(* IEC 61131-3 sources: STAR-PLC-Agent/results/raw/codex_matrix_resume_20261114/codex_deepseek/PUB011/functional/attempt_0001, 1 file *)

(* ---- test_program.st ---- *)
PROGRAM PLC_PRG
VAR
 BenchStep : UDINT := 0;
 BenchCalls : UDINT := 0;
 BenchDone : BOOL := FALSE;
 BenchUut0 : FB_Task;
 BenchUut1 : FB_Task;
 BenchUut2 : FB_Task;
 BenchUut3 : FB_Task;
 BenchUut4 : FB_Task;
 BenchUut5 : FB_Task;
 BenchUut6 : FB_Task;
 BenchUut7 : FB_Task;
 TraceIn_Mode : ARRAY[0..81] OF BOOL;
 TraceIn_ForwardButton : ARRAY[0..81] OF BOOL;
 TraceIn_ReverseButton : ARRAY[0..81] OF BOOL;
 TraceIn_SensorA : ARRAY[0..81] OF BOOL;
 TraceIn_SensorB : ARRAY[0..81] OF BOOL;
 TraceIn_SensorC : ARRAY[0..81] OF BOOL;
 TraceIn_ButtonA : ARRAY[0..81] OF BOOL;
 TraceIn_ButtonB : ARRAY[0..81] OF BOOL;
 TraceIn_ButtonC : ARRAY[0..81] OF BOOL;
 TraceOut_MotorForward : ARRAY[0..81] OF BOOL;
 TraceOut_MotorReverse : ARRAY[0..81] OF BOOL;
 TraceOut_CompletionLight : ARRAY[0..81] OF BOOL;
END_VAR

IF NOT BenchDone THEN
 CASE BenchStep OF
 0:
   BenchUut0.Mode := FALSE;
   BenchUut0.ForwardButton := FALSE;
   BenchUut0.ReverseButton := FALSE;
   BenchUut0.SensorA := FALSE;
   BenchUut0.SensorB := FALSE;
   BenchUut0.SensorC := FALSE;
   BenchUut0.ButtonA := FALSE;
   BenchUut0.ButtonB := FALSE;
   BenchUut0.ButtonC := FALSE;
   TraceIn_Mode[0] := BenchUut0.Mode;
   TraceIn_ForwardButton[0] := BenchUut0.ForwardButton;
   TraceIn_ReverseButton[0] := BenchUut0.ReverseButton;
   TraceIn_SensorA[0] := BenchUut0.SensorA;
   TraceIn_SensorB[0] := BenchUut0.SensorB;
   TraceIn_SensorC[0] := BenchUut0.SensorC;
   TraceIn_ButtonA[0] := BenchUut0.ButtonA;
   TraceIn_ButtonB[0] := BenchUut0.ButtonB;
   TraceIn_ButtonC[0] := BenchUut0.ButtonC;
   BenchUut0();
   TraceOut_MotorForward[0] := BenchUut0.MotorForward;
   TraceOut_MotorReverse[0] := BenchUut0.MotorReverse;
   TraceOut_CompletionLight[0] := BenchUut0.CompletionLight;
   BenchCalls := BenchCalls + 1;
 1:
   BenchUut0.Mode := FALSE;
   BenchUut0.ForwardButton := TRUE;
   BenchUut0.ReverseButton := FALSE;
   BenchUut0.SensorA := FALSE;
   BenchUut0.SensorB := FALSE;
   BenchUut0.SensorC := FALSE;
   BenchUut0.ButtonA := FALSE;
   BenchUut0.ButtonB := FALSE;
   BenchUut0.ButtonC := FALSE;
   TraceIn_Mode[1] := BenchUut0.Mode;
   TraceIn_ForwardButton[1] := BenchUut0.ForwardButton;
   TraceIn_ReverseButton[1] := BenchUut0.ReverseButton;
   TraceIn_SensorA[1] := BenchUut0.SensorA;
   TraceIn_SensorB[1] := BenchUut0.SensorB;
   TraceIn_SensorC[1] := BenchUut0.SensorC;
   TraceIn_ButtonA[1] := BenchUut0.ButtonA;
   TraceIn_ButtonB[1] := BenchUut0.ButtonB;
   TraceIn_ButtonC[1] := BenchUut0.ButtonC;
   BenchUut0();
   TraceOut_MotorForward[1] := BenchUut0.MotorForward;
   TraceOut_MotorReverse[1] := BenchUut0.MotorReverse;
   TraceOut_CompletionLight[1] := BenchUut0.CompletionLight;
   BenchCalls := BenchCalls + 1;
 2:
   BenchUut0.Mode := FALSE;
   BenchUut0.ForwardButton := FALSE;
   BenchUut0.ReverseButton := TRUE;
   BenchUut0.SensorA := FALSE;
   BenchUut0.SensorB := FALSE;
   BenchUut0.SensorC := FALSE;
   BenchUut0.ButtonA := FALSE;
   BenchUut0.ButtonB := FALSE;
   BenchUut0.ButtonC := FALSE;
   TraceIn_Mode[2] := BenchUut0.Mode;
   TraceIn_ForwardButton[2] := BenchUut0.ForwardButton;
   TraceIn_ReverseButton[2] := BenchUut0.ReverseButton;
   TraceIn_SensorA[2] := BenchUut0.SensorA;
   TraceIn_SensorB[2] := BenchUut0.SensorB;
   TraceIn_SensorC[2] := BenchUut0.SensorC;
   TraceIn_ButtonA[2] := BenchUut0.ButtonA;
   TraceIn_ButtonB[2] := BenchUut0.ButtonB;
   TraceIn_ButtonC[2] := BenchUut0.ButtonC;
   BenchUut0();
   TraceOut_MotorForward[2] := BenchUut0.MotorForward;
   TraceOut_MotorReverse[2] := BenchUut0.MotorReverse;
   TraceOut_CompletionLight[2] := BenchUut0.CompletionLight;
   BenchCalls := BenchCalls + 1;
 3:
   BenchUut1.Mode := TRUE;
   BenchUut1.ForwardButton := FALSE;
   BenchUut1.ReverseButton := FALSE;
   BenchUut1.SensorA := FALSE;
   BenchUut1.SensorB := FALSE;
   BenchUut1.SensorC := FALSE;
   BenchUut1.ButtonA := FALSE;
   BenchUut1.ButtonB := FALSE;
   BenchUut1.ButtonC := FALSE;
   TraceIn_Mode[3] := BenchUut1.Mode;
   TraceIn_ForwardButton[3] := BenchUut1.ForwardButton;
   TraceIn_ReverseButton[3] := BenchUut1.ReverseButton;
   TraceIn_SensorA[3] := BenchUut1.SensorA;
   TraceIn_SensorB[3] := BenchUut1.SensorB;
   TraceIn_SensorC[3] := BenchUut1.SensorC;
   TraceIn_ButtonA[3] := BenchUut1.ButtonA;
   TraceIn_ButtonB[3] := BenchUut1.ButtonB;
   TraceIn_ButtonC[3] := BenchUut1.ButtonC;
   BenchUut1();
   TraceOut_MotorForward[3] := BenchUut1.MotorForward;
   TraceOut_MotorReverse[3] := BenchUut1.MotorReverse;
   TraceOut_CompletionLight[3] := BenchUut1.CompletionLight;
   BenchCalls := BenchCalls + 1;
 4:
   BenchUut1.Mode := TRUE;
   BenchUut1.ForwardButton := FALSE;
   BenchUut1.ReverseButton := FALSE;
   BenchUut1.SensorA := TRUE;
   BenchUut1.SensorB := FALSE;
   BenchUut1.SensorC := FALSE;
   BenchUut1.ButtonA := FALSE;
   BenchUut1.ButtonB := FALSE;
   BenchUut1.ButtonC := FALSE;
   TraceIn_Mode[4] := BenchUut1.Mode;
   TraceIn_ForwardButton[4] := BenchUut1.ForwardButton;
   TraceIn_ReverseButton[4] := BenchUut1.ReverseButton;
   TraceIn_SensorA[4] := BenchUut1.SensorA;
   TraceIn_SensorB[4] := BenchUut1.SensorB;
   TraceIn_SensorC[4] := BenchUut1.SensorC;
   TraceIn_ButtonA[4] := BenchUut1.ButtonA;
   TraceIn_ButtonB[4] := BenchUut1.ButtonB;
   TraceIn_ButtonC[4] := BenchUut1.ButtonC;
   BenchUut1();
   TraceOut_MotorForward[4] := BenchUut1.MotorForward;
   TraceOut_MotorReverse[4] := BenchUut1.MotorReverse;
   TraceOut_CompletionLight[4] := BenchUut1.CompletionLight;
   BenchCalls := BenchCalls + 1;
 5:
   BenchUut1.Mode := TRUE;
   BenchUut1.ForwardButton := FALSE;
   BenchUut1.ReverseButton := FALSE;
   BenchUut1.SensorA := TRUE;
   BenchUut1.SensorB := FALSE;
   BenchUut1.SensorC := FALSE;
   BenchUut1.ButtonA := TRUE;
   BenchUut1.ButtonB := FALSE;
   BenchUut1.ButtonC := FALSE;
   TraceIn_Mode[5] := BenchUut1.Mode;
   TraceIn_ForwardButton[5] := BenchUut1.ForwardButton;
   TraceIn_ReverseButton[5] := BenchUut1.ReverseButton;
   TraceIn_SensorA[5] := BenchUut1.SensorA;
   TraceIn_SensorB[5] := BenchUut1.SensorB;
   TraceIn_SensorC[5] := BenchUut1.SensorC;
   TraceIn_ButtonA[5] := BenchUut1.ButtonA;
   TraceIn_ButtonB[5] := BenchUut1.ButtonB;
   TraceIn_ButtonC[5] := BenchUut1.ButtonC;
   BenchUut1();
   TraceOut_MotorForward[5] := BenchUut1.MotorForward;
   TraceOut_MotorReverse[5] := BenchUut1.MotorReverse;
   TraceOut_CompletionLight[5] := BenchUut1.CompletionLight;
   BenchCalls := BenchCalls + 1;
 6:
   BenchUut1.Mode := TRUE;
   BenchUut1.ForwardButton := FALSE;
   BenchUut1.ReverseButton := FALSE;
   BenchUut1.SensorA := FALSE;
   BenchUut1.SensorB := FALSE;
   BenchUut1.SensorC := FALSE;
   BenchUut1.ButtonA := FALSE;
   BenchUut1.ButtonB := FALSE;
   BenchUut1.ButtonC := FALSE;
   TraceIn_Mode[6] := BenchUut1.Mode;
   TraceIn_ForwardButton[6] := BenchUut1.ForwardButton;
   TraceIn_ReverseButton[6] := BenchUut1.ReverseButton;
   TraceIn_SensorA[6] := BenchUut1.SensorA;
   TraceIn_SensorB[6] := BenchUut1.SensorB;
   TraceIn_SensorC[6] := BenchUut1.SensorC;
   TraceIn_ButtonA[6] := BenchUut1.ButtonA;
   TraceIn_ButtonB[6] := BenchUut1.ButtonB;
   TraceIn_ButtonC[6] := BenchUut1.ButtonC;
   BenchUut1();
   TraceOut_MotorForward[6] := BenchUut1.MotorForward;
   TraceOut_MotorReverse[6] := BenchUut1.MotorReverse;
   TraceOut_CompletionLight[6] := BenchUut1.CompletionLight;
   BenchCalls := BenchCalls + 1;
 7:
   BenchUut1.Mode := TRUE;
   BenchUut1.ForwardButton := FALSE;
   BenchUut1.ReverseButton := FALSE;
   BenchUut1.SensorA := FALSE;
   BenchUut1.SensorB := TRUE;
   BenchUut1.SensorC := FALSE;
   BenchUut1.ButtonA := FALSE;
   BenchUut1.ButtonB := FALSE;
   BenchUut1.ButtonC := FALSE;
   TraceIn_Mode[7] := BenchUut1.Mode;
   TraceIn_ForwardButton[7] := BenchUut1.ForwardButton;
   TraceIn_ReverseButton[7] := BenchUut1.ReverseButton;
   TraceIn_SensorA[7] := BenchUut1.SensorA;
   TraceIn_SensorB[7] := BenchUut1.SensorB;
   TraceIn_SensorC[7] := BenchUut1.SensorC;
   TraceIn_ButtonA[7] := BenchUut1.ButtonA;
   TraceIn_ButtonB[7] := BenchUut1.ButtonB;
   TraceIn_ButtonC[7] := BenchUut1.ButtonC;
   BenchUut1();
   TraceOut_MotorForward[7] := BenchUut1.MotorForward;
   TraceOut_MotorReverse[7] := BenchUut1.MotorReverse;
   TraceOut_CompletionLight[7] := BenchUut1.CompletionLight;
   BenchCalls := BenchCalls + 1;
 8:
   BenchUut1.Mode := TRUE;
   BenchUut1.ForwardButton := FALSE;
   BenchUut1.ReverseButton := FALSE;
   BenchUut1.SensorA := FALSE;
   BenchUut1.SensorB := TRUE;
   BenchUut1.SensorC := FALSE;
   BenchUut1.ButtonA := FALSE;
   BenchUut1.ButtonB := TRUE;
   BenchUut1.ButtonC := FALSE;
   TraceIn_Mode[8] := BenchUut1.Mode;
   TraceIn_ForwardButton[8] := BenchUut1.ForwardButton;
   TraceIn_ReverseButton[8] := BenchUut1.ReverseButton;
   TraceIn_SensorA[8] := BenchUut1.SensorA;
   TraceIn_SensorB[8] := BenchUut1.SensorB;
   TraceIn_SensorC[8] := BenchUut1.SensorC;
   TraceIn_ButtonA[8] := BenchUut1.ButtonA;
   TraceIn_ButtonB[8] := BenchUut1.ButtonB;
   TraceIn_ButtonC[8] := BenchUut1.ButtonC;
   BenchUut1();
   TraceOut_MotorForward[8] := BenchUut1.MotorForward;
   TraceOut_MotorReverse[8] := BenchUut1.MotorReverse;
   TraceOut_CompletionLight[8] := BenchUut1.CompletionLight;
   BenchCalls := BenchCalls + 1;
 9:
   BenchUut1.Mode := TRUE;
   BenchUut1.ForwardButton := FALSE;
   BenchUut1.ReverseButton := FALSE;
   BenchUut1.SensorA := FALSE;
   BenchUut1.SensorB := FALSE;
   BenchUut1.SensorC := TRUE;
   BenchUut1.ButtonA := FALSE;
   BenchUut1.ButtonB := FALSE;
   BenchUut1.ButtonC := FALSE;
   TraceIn_Mode[9] := BenchUut1.Mode;
   TraceIn_ForwardButton[9] := BenchUut1.ForwardButton;
   TraceIn_ReverseButton[9] := BenchUut1.ReverseButton;
   TraceIn_SensorA[9] := BenchUut1.SensorA;
   TraceIn_SensorB[9] := BenchUut1.SensorB;
   TraceIn_SensorC[9] := BenchUut1.SensorC;
   TraceIn_ButtonA[9] := BenchUut1.ButtonA;
   TraceIn_ButtonB[9] := BenchUut1.ButtonB;
   TraceIn_ButtonC[9] := BenchUut1.ButtonC;
   BenchUut1();
   TraceOut_MotorForward[9] := BenchUut1.MotorForward;
   TraceOut_MotorReverse[9] := BenchUut1.MotorReverse;
   TraceOut_CompletionLight[9] := BenchUut1.CompletionLight;
   BenchCalls := BenchCalls + 1;
 10:
   BenchUut1.Mode := TRUE;
   BenchUut1.ForwardButton := FALSE;
   BenchUut1.ReverseButton := FALSE;
   BenchUut1.SensorA := FALSE;
   BenchUut1.SensorB := FALSE;
   BenchUut1.SensorC := TRUE;
   BenchUut1.ButtonA := FALSE;
   BenchUut1.ButtonB := FALSE;
   BenchUut1.ButtonC := TRUE;
   TraceIn_Mode[10] := BenchUut1.Mode;
   TraceIn_ForwardButton[10] := BenchUut1.ForwardButton;
   TraceIn_ReverseButton[10] := BenchUut1.ReverseButton;
   TraceIn_SensorA[10] := BenchUut1.SensorA;
   TraceIn_SensorB[10] := BenchUut1.SensorB;
   TraceIn_SensorC[10] := BenchUut1.SensorC;
   TraceIn_ButtonA[10] := BenchUut1.ButtonA;
   TraceIn_ButtonB[10] := BenchUut1.ButtonB;
   TraceIn_ButtonC[10] := BenchUut1.ButtonC;
   BenchUut1();
   TraceOut_MotorForward[10] := BenchUut1.MotorForward;
   TraceOut_MotorReverse[10] := BenchUut1.MotorReverse;
   TraceOut_CompletionLight[10] := BenchUut1.CompletionLight;
   BenchCalls := BenchCalls + 1;
 11:
   BenchUut1.Mode := TRUE;
   BenchUut1.ForwardButton := FALSE;
   BenchUut1.ReverseButton := FALSE;
   BenchUut1.SensorA := FALSE;
   BenchUut1.SensorB := FALSE;
   BenchUut1.SensorC := TRUE;
   BenchUut1.ButtonA := FALSE;
   BenchUut1.ButtonB := FALSE;
   BenchUut1.ButtonC := FALSE;
   TraceIn_Mode[11] := BenchUut1.Mode;
   TraceIn_ForwardButton[11] := BenchUut1.ForwardButton;
   TraceIn_ReverseButton[11] := BenchUut1.ReverseButton;
   TraceIn_SensorA[11] := BenchUut1.SensorA;
   TraceIn_SensorB[11] := BenchUut1.SensorB;
   TraceIn_SensorC[11] := BenchUut1.SensorC;
   TraceIn_ButtonA[11] := BenchUut1.ButtonA;
   TraceIn_ButtonB[11] := BenchUut1.ButtonB;
   TraceIn_ButtonC[11] := BenchUut1.ButtonC;
   BenchUut1();
   TraceOut_MotorForward[11] := BenchUut1.MotorForward;
   TraceOut_MotorReverse[11] := BenchUut1.MotorReverse;
   TraceOut_CompletionLight[11] := BenchUut1.CompletionLight;
   BenchCalls := BenchCalls + 1;
 12:
   BenchUut1.Mode := TRUE;
   BenchUut1.ForwardButton := FALSE;
   BenchUut1.ReverseButton := FALSE;
   BenchUut1.SensorA := FALSE;
   BenchUut1.SensorB := FALSE;
   BenchUut1.SensorC := FALSE;
   BenchUut1.ButtonA := FALSE;
   BenchUut1.ButtonB := FALSE;
   BenchUut1.ButtonC := FALSE;
   TraceIn_Mode[12] := BenchUut1.Mode;
   TraceIn_ForwardButton[12] := BenchUut1.ForwardButton;
   TraceIn_ReverseButton[12] := BenchUut1.ReverseButton;
   TraceIn_SensorA[12] := BenchUut1.SensorA;
   TraceIn_SensorB[12] := BenchUut1.SensorB;
   TraceIn_SensorC[12] := BenchUut1.SensorC;
   TraceIn_ButtonA[12] := BenchUut1.ButtonA;
   TraceIn_ButtonB[12] := BenchUut1.ButtonB;
   TraceIn_ButtonC[12] := BenchUut1.ButtonC;
   BenchUut1();
   TraceOut_MotorForward[12] := BenchUut1.MotorForward;
   TraceOut_MotorReverse[12] := BenchUut1.MotorReverse;
   TraceOut_CompletionLight[12] := BenchUut1.CompletionLight;
   BenchCalls := BenchCalls + 1;
 13:
   BenchUut2.Mode := TRUE;
   BenchUut2.ForwardButton := FALSE;
   BenchUut2.ReverseButton := FALSE;
   BenchUut2.SensorA := FALSE;
   BenchUut2.SensorB := FALSE;
   BenchUut2.SensorC := FALSE;
   BenchUut2.ButtonA := FALSE;
   BenchUut2.ButtonB := TRUE;
   BenchUut2.ButtonC := TRUE;
   TraceIn_Mode[13] := BenchUut2.Mode;
   TraceIn_ForwardButton[13] := BenchUut2.ForwardButton;
   TraceIn_ReverseButton[13] := BenchUut2.ReverseButton;
   TraceIn_SensorA[13] := BenchUut2.SensorA;
   TraceIn_SensorB[13] := BenchUut2.SensorB;
   TraceIn_SensorC[13] := BenchUut2.SensorC;
   TraceIn_ButtonA[13] := BenchUut2.ButtonA;
   TraceIn_ButtonB[13] := BenchUut2.ButtonB;
   TraceIn_ButtonC[13] := BenchUut2.ButtonC;
   BenchUut2();
   TraceOut_MotorForward[13] := BenchUut2.MotorForward;
   TraceOut_MotorReverse[13] := BenchUut2.MotorReverse;
   TraceOut_CompletionLight[13] := BenchUut2.CompletionLight;
   BenchCalls := BenchCalls + 1;
 14:
   BenchUut2.Mode := TRUE;
   BenchUut2.ForwardButton := FALSE;
   BenchUut2.ReverseButton := FALSE;
   BenchUut2.SensorA := TRUE;
   BenchUut2.SensorB := FALSE;
   BenchUut2.SensorC := FALSE;
   BenchUut2.ButtonA := FALSE;
   BenchUut2.ButtonB := TRUE;
   BenchUut2.ButtonC := FALSE;
   TraceIn_Mode[14] := BenchUut2.Mode;
   TraceIn_ForwardButton[14] := BenchUut2.ForwardButton;
   TraceIn_ReverseButton[14] := BenchUut2.ReverseButton;
   TraceIn_SensorA[14] := BenchUut2.SensorA;
   TraceIn_SensorB[14] := BenchUut2.SensorB;
   TraceIn_SensorC[14] := BenchUut2.SensorC;
   TraceIn_ButtonA[14] := BenchUut2.ButtonA;
   TraceIn_ButtonB[14] := BenchUut2.ButtonB;
   TraceIn_ButtonC[14] := BenchUut2.ButtonC;
   BenchUut2();
   TraceOut_MotorForward[14] := BenchUut2.MotorForward;
   TraceOut_MotorReverse[14] := BenchUut2.MotorReverse;
   TraceOut_CompletionLight[14] := BenchUut2.CompletionLight;
   BenchCalls := BenchCalls + 1;
 15:
   BenchUut3.Mode := TRUE;
   BenchUut3.ForwardButton := FALSE;
   BenchUut3.ReverseButton := FALSE;
   BenchUut3.SensorA := FALSE;
   BenchUut3.SensorB := FALSE;
   BenchUut3.SensorC := FALSE;
   BenchUut3.ButtonA := FALSE;
   BenchUut3.ButtonB := FALSE;
   BenchUut3.ButtonC := FALSE;
   TraceIn_Mode[15] := BenchUut3.Mode;
   TraceIn_ForwardButton[15] := BenchUut3.ForwardButton;
   TraceIn_ReverseButton[15] := BenchUut3.ReverseButton;
   TraceIn_SensorA[15] := BenchUut3.SensorA;
   TraceIn_SensorB[15] := BenchUut3.SensorB;
   TraceIn_SensorC[15] := BenchUut3.SensorC;
   TraceIn_ButtonA[15] := BenchUut3.ButtonA;
   TraceIn_ButtonB[15] := BenchUut3.ButtonB;
   TraceIn_ButtonC[15] := BenchUut3.ButtonC;
   BenchUut3();
   TraceOut_MotorForward[15] := BenchUut3.MotorForward;
   TraceOut_MotorReverse[15] := BenchUut3.MotorReverse;
   TraceOut_CompletionLight[15] := BenchUut3.CompletionLight;
   BenchCalls := BenchCalls + 1;
 16:
   BenchUut3.Mode := TRUE;
   BenchUut3.ForwardButton := FALSE;
   BenchUut3.ReverseButton := FALSE;
   BenchUut3.SensorA := TRUE;
   BenchUut3.SensorB := FALSE;
   BenchUut3.SensorC := FALSE;
   BenchUut3.ButtonA := FALSE;
   BenchUut3.ButtonB := FALSE;
   BenchUut3.ButtonC := FALSE;
   TraceIn_Mode[16] := BenchUut3.Mode;
   TraceIn_ForwardButton[16] := BenchUut3.ForwardButton;
   TraceIn_ReverseButton[16] := BenchUut3.ReverseButton;
   TraceIn_SensorA[16] := BenchUut3.SensorA;
   TraceIn_SensorB[16] := BenchUut3.SensorB;
   TraceIn_SensorC[16] := BenchUut3.SensorC;
   TraceIn_ButtonA[16] := BenchUut3.ButtonA;
   TraceIn_ButtonB[16] := BenchUut3.ButtonB;
   TraceIn_ButtonC[16] := BenchUut3.ButtonC;
   BenchUut3();
   TraceOut_MotorForward[16] := BenchUut3.MotorForward;
   TraceOut_MotorReverse[16] := BenchUut3.MotorReverse;
   TraceOut_CompletionLight[16] := BenchUut3.CompletionLight;
   BenchCalls := BenchCalls + 1;
 17:
   BenchUut3.Mode := TRUE;
   BenchUut3.ForwardButton := FALSE;
   BenchUut3.ReverseButton := FALSE;
   BenchUut3.SensorA := TRUE;
   BenchUut3.SensorB := FALSE;
   BenchUut3.SensorC := FALSE;
   BenchUut3.ButtonA := TRUE;
   BenchUut3.ButtonB := FALSE;
   BenchUut3.ButtonC := FALSE;
   TraceIn_Mode[17] := BenchUut3.Mode;
   TraceIn_ForwardButton[17] := BenchUut3.ForwardButton;
   TraceIn_ReverseButton[17] := BenchUut3.ReverseButton;
   TraceIn_SensorA[17] := BenchUut3.SensorA;
   TraceIn_SensorB[17] := BenchUut3.SensorB;
   TraceIn_SensorC[17] := BenchUut3.SensorC;
   TraceIn_ButtonA[17] := BenchUut3.ButtonA;
   TraceIn_ButtonB[17] := BenchUut3.ButtonB;
   TraceIn_ButtonC[17] := BenchUut3.ButtonC;
   BenchUut3();
   TraceOut_MotorForward[17] := BenchUut3.MotorForward;
   TraceOut_MotorReverse[17] := BenchUut3.MotorReverse;
   TraceOut_CompletionLight[17] := BenchUut3.CompletionLight;
   BenchCalls := BenchCalls + 1;
 18:
   BenchUut3.Mode := TRUE;
   BenchUut3.ForwardButton := FALSE;
   BenchUut3.ReverseButton := FALSE;
   BenchUut3.SensorA := FALSE;
   BenchUut3.SensorB := FALSE;
   BenchUut3.SensorC := FALSE;
   BenchUut3.ButtonA := FALSE;
   BenchUut3.ButtonB := FALSE;
   BenchUut3.ButtonC := FALSE;
   TraceIn_Mode[18] := BenchUut3.Mode;
   TraceIn_ForwardButton[18] := BenchUut3.ForwardButton;
   TraceIn_ReverseButton[18] := BenchUut3.ReverseButton;
   TraceIn_SensorA[18] := BenchUut3.SensorA;
   TraceIn_SensorB[18] := BenchUut3.SensorB;
   TraceIn_SensorC[18] := BenchUut3.SensorC;
   TraceIn_ButtonA[18] := BenchUut3.ButtonA;
   TraceIn_ButtonB[18] := BenchUut3.ButtonB;
   TraceIn_ButtonC[18] := BenchUut3.ButtonC;
   BenchUut3();
   TraceOut_MotorForward[18] := BenchUut3.MotorForward;
   TraceOut_MotorReverse[18] := BenchUut3.MotorReverse;
   TraceOut_CompletionLight[18] := BenchUut3.CompletionLight;
   BenchCalls := BenchCalls + 1;
 19:
   BenchUut3.Mode := TRUE;
   BenchUut3.ForwardButton := FALSE;
   BenchUut3.ReverseButton := FALSE;
   BenchUut3.SensorA := FALSE;
   BenchUut3.SensorB := TRUE;
   BenchUut3.SensorC := FALSE;
   BenchUut3.ButtonA := FALSE;
   BenchUut3.ButtonB := FALSE;
   BenchUut3.ButtonC := FALSE;
   TraceIn_Mode[19] := BenchUut3.Mode;
   TraceIn_ForwardButton[19] := BenchUut3.ForwardButton;
   TraceIn_ReverseButton[19] := BenchUut3.ReverseButton;
   TraceIn_SensorA[19] := BenchUut3.SensorA;
   TraceIn_SensorB[19] := BenchUut3.SensorB;
   TraceIn_SensorC[19] := BenchUut3.SensorC;
   TraceIn_ButtonA[19] := BenchUut3.ButtonA;
   TraceIn_ButtonB[19] := BenchUut3.ButtonB;
   TraceIn_ButtonC[19] := BenchUut3.ButtonC;
   BenchUut3();
   TraceOut_MotorForward[19] := BenchUut3.MotorForward;
   TraceOut_MotorReverse[19] := BenchUut3.MotorReverse;
   TraceOut_CompletionLight[19] := BenchUut3.CompletionLight;
   BenchCalls := BenchCalls + 1;
 20:
   BenchUut3.Mode := TRUE;
   BenchUut3.ForwardButton := FALSE;
   BenchUut3.ReverseButton := FALSE;
   BenchUut3.SensorA := FALSE;
   BenchUut3.SensorB := TRUE;
   BenchUut3.SensorC := FALSE;
   BenchUut3.ButtonA := FALSE;
   BenchUut3.ButtonB := TRUE;
   BenchUut3.ButtonC := FALSE;
   TraceIn_Mode[20] := BenchUut3.Mode;
   TraceIn_ForwardButton[20] := BenchUut3.ForwardButton;
   TraceIn_ReverseButton[20] := BenchUut3.ReverseButton;
   TraceIn_SensorA[20] := BenchUut3.SensorA;
   TraceIn_SensorB[20] := BenchUut3.SensorB;
   TraceIn_SensorC[20] := BenchUut3.SensorC;
   TraceIn_ButtonA[20] := BenchUut3.ButtonA;
   TraceIn_ButtonB[20] := BenchUut3.ButtonB;
   TraceIn_ButtonC[20] := BenchUut3.ButtonC;
   BenchUut3();
   TraceOut_MotorForward[20] := BenchUut3.MotorForward;
   TraceOut_MotorReverse[20] := BenchUut3.MotorReverse;
   TraceOut_CompletionLight[20] := BenchUut3.CompletionLight;
   BenchCalls := BenchCalls + 1;
 21:
   BenchUut3.Mode := TRUE;
   BenchUut3.ForwardButton := FALSE;
   BenchUut3.ReverseButton := FALSE;
   BenchUut3.SensorA := FALSE;
   BenchUut3.SensorB := FALSE;
   BenchUut3.SensorC := FALSE;
   BenchUut3.ButtonA := FALSE;
   BenchUut3.ButtonB := FALSE;
   BenchUut3.ButtonC := FALSE;
   TraceIn_Mode[21] := BenchUut3.Mode;
   TraceIn_ForwardButton[21] := BenchUut3.ForwardButton;
   TraceIn_ReverseButton[21] := BenchUut3.ReverseButton;
   TraceIn_SensorA[21] := BenchUut3.SensorA;
   TraceIn_SensorB[21] := BenchUut3.SensorB;
   TraceIn_SensorC[21] := BenchUut3.SensorC;
   TraceIn_ButtonA[21] := BenchUut3.ButtonA;
   TraceIn_ButtonB[21] := BenchUut3.ButtonB;
   TraceIn_ButtonC[21] := BenchUut3.ButtonC;
   BenchUut3();
   TraceOut_MotorForward[21] := BenchUut3.MotorForward;
   TraceOut_MotorReverse[21] := BenchUut3.MotorReverse;
   TraceOut_CompletionLight[21] := BenchUut3.CompletionLight;
   BenchCalls := BenchCalls + 1;
 22:
   BenchUut4.Mode := TRUE;
   BenchUut4.ForwardButton := FALSE;
   BenchUut4.ReverseButton := FALSE;
   BenchUut4.SensorA := TRUE;
   BenchUut4.SensorB := FALSE;
   BenchUut4.SensorC := FALSE;
   BenchUut4.ButtonA := TRUE;
   BenchUut4.ButtonB := FALSE;
   BenchUut4.ButtonC := FALSE;
   TraceIn_Mode[22] := BenchUut4.Mode;
   TraceIn_ForwardButton[22] := BenchUut4.ForwardButton;
   TraceIn_ReverseButton[22] := BenchUut4.ReverseButton;
   TraceIn_SensorA[22] := BenchUut4.SensorA;
   TraceIn_SensorB[22] := BenchUut4.SensorB;
   TraceIn_SensorC[22] := BenchUut4.SensorC;
   TraceIn_ButtonA[22] := BenchUut4.ButtonA;
   TraceIn_ButtonB[22] := BenchUut4.ButtonB;
   TraceIn_ButtonC[22] := BenchUut4.ButtonC;
   BenchUut4();
   TraceOut_MotorForward[22] := BenchUut4.MotorForward;
   TraceOut_MotorReverse[22] := BenchUut4.MotorReverse;
   TraceOut_CompletionLight[22] := BenchUut4.CompletionLight;
   BenchCalls := BenchCalls + 1;
 23:
   BenchUut4.Mode := TRUE;
   BenchUut4.ForwardButton := FALSE;
   BenchUut4.ReverseButton := FALSE;
   BenchUut4.SensorA := FALSE;
   BenchUut4.SensorB := FALSE;
   BenchUut4.SensorC := FALSE;
   BenchUut4.ButtonA := FALSE;
   BenchUut4.ButtonB := FALSE;
   BenchUut4.ButtonC := FALSE;
   TraceIn_Mode[23] := BenchUut4.Mode;
   TraceIn_ForwardButton[23] := BenchUut4.ForwardButton;
   TraceIn_ReverseButton[23] := BenchUut4.ReverseButton;
   TraceIn_SensorA[23] := BenchUut4.SensorA;
   TraceIn_SensorB[23] := BenchUut4.SensorB;
   TraceIn_SensorC[23] := BenchUut4.SensorC;
   TraceIn_ButtonA[23] := BenchUut4.ButtonA;
   TraceIn_ButtonB[23] := BenchUut4.ButtonB;
   TraceIn_ButtonC[23] := BenchUut4.ButtonC;
   BenchUut4();
   TraceOut_MotorForward[23] := BenchUut4.MotorForward;
   TraceOut_MotorReverse[23] := BenchUut4.MotorReverse;
   TraceOut_CompletionLight[23] := BenchUut4.CompletionLight;
   BenchCalls := BenchCalls + 1;
 24:
   BenchUut4.Mode := FALSE;
   BenchUut4.ForwardButton := FALSE;
   BenchUut4.ReverseButton := TRUE;
   BenchUut4.SensorA := FALSE;
   BenchUut4.SensorB := FALSE;
   BenchUut4.SensorC := FALSE;
   BenchUut4.ButtonA := FALSE;
   BenchUut4.ButtonB := FALSE;
   BenchUut4.ButtonC := FALSE;
   TraceIn_Mode[24] := BenchUut4.Mode;
   TraceIn_ForwardButton[24] := BenchUut4.ForwardButton;
   TraceIn_ReverseButton[24] := BenchUut4.ReverseButton;
   TraceIn_SensorA[24] := BenchUut4.SensorA;
   TraceIn_SensorB[24] := BenchUut4.SensorB;
   TraceIn_SensorC[24] := BenchUut4.SensorC;
   TraceIn_ButtonA[24] := BenchUut4.ButtonA;
   TraceIn_ButtonB[24] := BenchUut4.ButtonB;
   TraceIn_ButtonC[24] := BenchUut4.ButtonC;
   BenchUut4();
   TraceOut_MotorForward[24] := BenchUut4.MotorForward;
   TraceOut_MotorReverse[24] := BenchUut4.MotorReverse;
   TraceOut_CompletionLight[24] := BenchUut4.CompletionLight;
   BenchCalls := BenchCalls + 1;
 25:
   BenchUut4.Mode := TRUE;
   BenchUut4.ForwardButton := FALSE;
   BenchUut4.ReverseButton := FALSE;
   BenchUut4.SensorA := FALSE;
   BenchUut4.SensorB := FALSE;
   BenchUut4.SensorC := FALSE;
   BenchUut4.ButtonA := FALSE;
   BenchUut4.ButtonB := FALSE;
   BenchUut4.ButtonC := FALSE;
   TraceIn_Mode[25] := BenchUut4.Mode;
   TraceIn_ForwardButton[25] := BenchUut4.ForwardButton;
   TraceIn_ReverseButton[25] := BenchUut4.ReverseButton;
   TraceIn_SensorA[25] := BenchUut4.SensorA;
   TraceIn_SensorB[25] := BenchUut4.SensorB;
   TraceIn_SensorC[25] := BenchUut4.SensorC;
   TraceIn_ButtonA[25] := BenchUut4.ButtonA;
   TraceIn_ButtonB[25] := BenchUut4.ButtonB;
   TraceIn_ButtonC[25] := BenchUut4.ButtonC;
   BenchUut4();
   TraceOut_MotorForward[25] := BenchUut4.MotorForward;
   TraceOut_MotorReverse[25] := BenchUut4.MotorReverse;
   TraceOut_CompletionLight[25] := BenchUut4.CompletionLight;
   BenchCalls := BenchCalls + 1;
 26:
   BenchUut4.Mode := TRUE;
   BenchUut4.ForwardButton := FALSE;
   BenchUut4.ReverseButton := FALSE;
   BenchUut4.SensorA := TRUE;
   BenchUut4.SensorB := FALSE;
   BenchUut4.SensorC := FALSE;
   BenchUut4.ButtonA := FALSE;
   BenchUut4.ButtonB := FALSE;
   BenchUut4.ButtonC := FALSE;
   TraceIn_Mode[26] := BenchUut4.Mode;
   TraceIn_ForwardButton[26] := BenchUut4.ForwardButton;
   TraceIn_ReverseButton[26] := BenchUut4.ReverseButton;
   TraceIn_SensorA[26] := BenchUut4.SensorA;
   TraceIn_SensorB[26] := BenchUut4.SensorB;
   TraceIn_SensorC[26] := BenchUut4.SensorC;
   TraceIn_ButtonA[26] := BenchUut4.ButtonA;
   TraceIn_ButtonB[26] := BenchUut4.ButtonB;
   TraceIn_ButtonC[26] := BenchUut4.ButtonC;
   BenchUut4();
   TraceOut_MotorForward[26] := BenchUut4.MotorForward;
   TraceOut_MotorReverse[26] := BenchUut4.MotorReverse;
   TraceOut_CompletionLight[26] := BenchUut4.CompletionLight;
   BenchCalls := BenchCalls + 1;
 27:
   BenchUut4.Mode := TRUE;
   BenchUut4.ForwardButton := FALSE;
   BenchUut4.ReverseButton := FALSE;
   BenchUut4.SensorA := TRUE;
   BenchUut4.SensorB := FALSE;
   BenchUut4.SensorC := FALSE;
   BenchUut4.ButtonA := TRUE;
   BenchUut4.ButtonB := FALSE;
   BenchUut4.ButtonC := FALSE;
   TraceIn_Mode[27] := BenchUut4.Mode;
   TraceIn_ForwardButton[27] := BenchUut4.ForwardButton;
   TraceIn_ReverseButton[27] := BenchUut4.ReverseButton;
   TraceIn_SensorA[27] := BenchUut4.SensorA;
   TraceIn_SensorB[27] := BenchUut4.SensorB;
   TraceIn_SensorC[27] := BenchUut4.SensorC;
   TraceIn_ButtonA[27] := BenchUut4.ButtonA;
   TraceIn_ButtonB[27] := BenchUut4.ButtonB;
   TraceIn_ButtonC[27] := BenchUut4.ButtonC;
   BenchUut4();
   TraceOut_MotorForward[27] := BenchUut4.MotorForward;
   TraceOut_MotorReverse[27] := BenchUut4.MotorReverse;
   TraceOut_CompletionLight[27] := BenchUut4.CompletionLight;
   BenchCalls := BenchCalls + 1;
 28:
   BenchUut4.Mode := TRUE;
   BenchUut4.ForwardButton := FALSE;
   BenchUut4.ReverseButton := FALSE;
   BenchUut4.SensorA := FALSE;
   BenchUut4.SensorB := TRUE;
   BenchUut4.SensorC := FALSE;
   BenchUut4.ButtonA := FALSE;
   BenchUut4.ButtonB := TRUE;
   BenchUut4.ButtonC := FALSE;
   TraceIn_Mode[28] := BenchUut4.Mode;
   TraceIn_ForwardButton[28] := BenchUut4.ForwardButton;
   TraceIn_ReverseButton[28] := BenchUut4.ReverseButton;
   TraceIn_SensorA[28] := BenchUut4.SensorA;
   TraceIn_SensorB[28] := BenchUut4.SensorB;
   TraceIn_SensorC[28] := BenchUut4.SensorC;
   TraceIn_ButtonA[28] := BenchUut4.ButtonA;
   TraceIn_ButtonB[28] := BenchUut4.ButtonB;
   TraceIn_ButtonC[28] := BenchUut4.ButtonC;
   BenchUut4();
   TraceOut_MotorForward[28] := BenchUut4.MotorForward;
   TraceOut_MotorReverse[28] := BenchUut4.MotorReverse;
   TraceOut_CompletionLight[28] := BenchUut4.CompletionLight;
   BenchCalls := BenchCalls + 1;
 29:
   BenchUut4.Mode := TRUE;
   BenchUut4.ForwardButton := FALSE;
   BenchUut4.ReverseButton := FALSE;
   BenchUut4.SensorA := FALSE;
   BenchUut4.SensorB := TRUE;
   BenchUut4.SensorC := FALSE;
   BenchUut4.ButtonA := FALSE;
   BenchUut4.ButtonB := FALSE;
   BenchUut4.ButtonC := FALSE;
   TraceIn_Mode[29] := BenchUut4.Mode;
   TraceIn_ForwardButton[29] := BenchUut4.ForwardButton;
   TraceIn_ReverseButton[29] := BenchUut4.ReverseButton;
   TraceIn_SensorA[29] := BenchUut4.SensorA;
   TraceIn_SensorB[29] := BenchUut4.SensorB;
   TraceIn_SensorC[29] := BenchUut4.SensorC;
   TraceIn_ButtonA[29] := BenchUut4.ButtonA;
   TraceIn_ButtonB[29] := BenchUut4.ButtonB;
   TraceIn_ButtonC[29] := BenchUut4.ButtonC;
   BenchUut4();
   TraceOut_MotorForward[29] := BenchUut4.MotorForward;
   TraceOut_MotorReverse[29] := BenchUut4.MotorReverse;
   TraceOut_CompletionLight[29] := BenchUut4.CompletionLight;
   BenchCalls := BenchCalls + 1;
 30:
   BenchUut4.Mode := TRUE;
   BenchUut4.ForwardButton := FALSE;
   BenchUut4.ReverseButton := FALSE;
   BenchUut4.SensorA := FALSE;
   BenchUut4.SensorB := TRUE;
   BenchUut4.SensorC := FALSE;
   BenchUut4.ButtonA := FALSE;
   BenchUut4.ButtonB := TRUE;
   BenchUut4.ButtonC := FALSE;
   TraceIn_Mode[30] := BenchUut4.Mode;
   TraceIn_ForwardButton[30] := BenchUut4.ForwardButton;
   TraceIn_ReverseButton[30] := BenchUut4.ReverseButton;
   TraceIn_SensorA[30] := BenchUut4.SensorA;
   TraceIn_SensorB[30] := BenchUut4.SensorB;
   TraceIn_SensorC[30] := BenchUut4.SensorC;
   TraceIn_ButtonA[30] := BenchUut4.ButtonA;
   TraceIn_ButtonB[30] := BenchUut4.ButtonB;
   TraceIn_ButtonC[30] := BenchUut4.ButtonC;
   BenchUut4();
   TraceOut_MotorForward[30] := BenchUut4.MotorForward;
   TraceOut_MotorReverse[30] := BenchUut4.MotorReverse;
   TraceOut_CompletionLight[30] := BenchUut4.CompletionLight;
   BenchCalls := BenchCalls + 1;
 31:
   BenchUut4.Mode := TRUE;
   BenchUut4.ForwardButton := FALSE;
   BenchUut4.ReverseButton := FALSE;
   BenchUut4.SensorA := FALSE;
   BenchUut4.SensorB := FALSE;
   BenchUut4.SensorC := TRUE;
   BenchUut4.ButtonA := FALSE;
   BenchUut4.ButtonB := FALSE;
   BenchUut4.ButtonC := TRUE;
   TraceIn_Mode[31] := BenchUut4.Mode;
   TraceIn_ForwardButton[31] := BenchUut4.ForwardButton;
   TraceIn_ReverseButton[31] := BenchUut4.ReverseButton;
   TraceIn_SensorA[31] := BenchUut4.SensorA;
   TraceIn_SensorB[31] := BenchUut4.SensorB;
   TraceIn_SensorC[31] := BenchUut4.SensorC;
   TraceIn_ButtonA[31] := BenchUut4.ButtonA;
   TraceIn_ButtonB[31] := BenchUut4.ButtonB;
   TraceIn_ButtonC[31] := BenchUut4.ButtonC;
   BenchUut4();
   TraceOut_MotorForward[31] := BenchUut4.MotorForward;
   TraceOut_MotorReverse[31] := BenchUut4.MotorReverse;
   TraceOut_CompletionLight[31] := BenchUut4.CompletionLight;
   BenchCalls := BenchCalls + 1;
 32:
   BenchUut4.Mode := TRUE;
   BenchUut4.ForwardButton := FALSE;
   BenchUut4.ReverseButton := FALSE;
   BenchUut4.SensorA := FALSE;
   BenchUut4.SensorB := FALSE;
   BenchUut4.SensorC := TRUE;
   BenchUut4.ButtonA := FALSE;
   BenchUut4.ButtonB := FALSE;
   BenchUut4.ButtonC := TRUE;
   TraceIn_Mode[32] := BenchUut4.Mode;
   TraceIn_ForwardButton[32] := BenchUut4.ForwardButton;
   TraceIn_ReverseButton[32] := BenchUut4.ReverseButton;
   TraceIn_SensorA[32] := BenchUut4.SensorA;
   TraceIn_SensorB[32] := BenchUut4.SensorB;
   TraceIn_SensorC[32] := BenchUut4.SensorC;
   TraceIn_ButtonA[32] := BenchUut4.ButtonA;
   TraceIn_ButtonB[32] := BenchUut4.ButtonB;
   TraceIn_ButtonC[32] := BenchUut4.ButtonC;
   BenchUut4();
   TraceOut_MotorForward[32] := BenchUut4.MotorForward;
   TraceOut_MotorReverse[32] := BenchUut4.MotorReverse;
   TraceOut_CompletionLight[32] := BenchUut4.CompletionLight;
   BenchCalls := BenchCalls + 1;
 33:
   BenchUut4.Mode := TRUE;
   BenchUut4.ForwardButton := FALSE;
   BenchUut4.ReverseButton := FALSE;
   BenchUut4.SensorA := FALSE;
   BenchUut4.SensorB := FALSE;
   BenchUut4.SensorC := FALSE;
   BenchUut4.ButtonA := FALSE;
   BenchUut4.ButtonB := FALSE;
   BenchUut4.ButtonC := FALSE;
   TraceIn_Mode[33] := BenchUut4.Mode;
   TraceIn_ForwardButton[33] := BenchUut4.ForwardButton;
   TraceIn_ReverseButton[33] := BenchUut4.ReverseButton;
   TraceIn_SensorA[33] := BenchUut4.SensorA;
   TraceIn_SensorB[33] := BenchUut4.SensorB;
   TraceIn_SensorC[33] := BenchUut4.SensorC;
   TraceIn_ButtonA[33] := BenchUut4.ButtonA;
   TraceIn_ButtonB[33] := BenchUut4.ButtonB;
   TraceIn_ButtonC[33] := BenchUut4.ButtonC;
   BenchUut4();
   TraceOut_MotorForward[33] := BenchUut4.MotorForward;
   TraceOut_MotorReverse[33] := BenchUut4.MotorReverse;
   TraceOut_CompletionLight[33] := BenchUut4.CompletionLight;
   BenchCalls := BenchCalls + 1;
 34:
   BenchUut5.Mode := FALSE;
   BenchUut5.ForwardButton := FALSE;
   BenchUut5.ReverseButton := FALSE;
   BenchUut5.SensorA := FALSE;
   BenchUut5.SensorB := FALSE;
   BenchUut5.SensorC := FALSE;
   BenchUut5.ButtonA := FALSE;
   BenchUut5.ButtonB := FALSE;
   BenchUut5.ButtonC := FALSE;
   TraceIn_Mode[34] := BenchUut5.Mode;
   TraceIn_ForwardButton[34] := BenchUut5.ForwardButton;
   TraceIn_ReverseButton[34] := BenchUut5.ReverseButton;
   TraceIn_SensorA[34] := BenchUut5.SensorA;
   TraceIn_SensorB[34] := BenchUut5.SensorB;
   TraceIn_SensorC[34] := BenchUut5.SensorC;
   TraceIn_ButtonA[34] := BenchUut5.ButtonA;
   TraceIn_ButtonB[34] := BenchUut5.ButtonB;
   TraceIn_ButtonC[34] := BenchUut5.ButtonC;
   BenchUut5();
   TraceOut_MotorForward[34] := BenchUut5.MotorForward;
   TraceOut_MotorReverse[34] := BenchUut5.MotorReverse;
   TraceOut_CompletionLight[34] := BenchUut5.CompletionLight;
   BenchCalls := BenchCalls + 1;
 35:
   BenchUut5.Mode := FALSE;
   BenchUut5.ForwardButton := FALSE;
   BenchUut5.ReverseButton := FALSE;
   BenchUut5.SensorA := FALSE;
   BenchUut5.SensorB := FALSE;
   BenchUut5.SensorC := FALSE;
   BenchUut5.ButtonA := FALSE;
   BenchUut5.ButtonB := FALSE;
   BenchUut5.ButtonC := FALSE;
   TraceIn_Mode[35] := BenchUut5.Mode;
   TraceIn_ForwardButton[35] := BenchUut5.ForwardButton;
   TraceIn_ReverseButton[35] := BenchUut5.ReverseButton;
   TraceIn_SensorA[35] := BenchUut5.SensorA;
   TraceIn_SensorB[35] := BenchUut5.SensorB;
   TraceIn_SensorC[35] := BenchUut5.SensorC;
   TraceIn_ButtonA[35] := BenchUut5.ButtonA;
   TraceIn_ButtonB[35] := BenchUut5.ButtonB;
   TraceIn_ButtonC[35] := BenchUut5.ButtonC;
   BenchUut5();
   TraceOut_MotorForward[35] := BenchUut5.MotorForward;
   TraceOut_MotorReverse[35] := BenchUut5.MotorReverse;
   TraceOut_CompletionLight[35] := BenchUut5.CompletionLight;
   BenchCalls := BenchCalls + 1;
 36:
   BenchUut5.Mode := FALSE;
   BenchUut5.ForwardButton := FALSE;
   BenchUut5.ReverseButton := FALSE;
   BenchUut5.SensorA := FALSE;
   BenchUut5.SensorB := FALSE;
   BenchUut5.SensorC := FALSE;
   BenchUut5.ButtonA := FALSE;
   BenchUut5.ButtonB := FALSE;
   BenchUut5.ButtonC := FALSE;
   TraceIn_Mode[36] := BenchUut5.Mode;
   TraceIn_ForwardButton[36] := BenchUut5.ForwardButton;
   TraceIn_ReverseButton[36] := BenchUut5.ReverseButton;
   TraceIn_SensorA[36] := BenchUut5.SensorA;
   TraceIn_SensorB[36] := BenchUut5.SensorB;
   TraceIn_SensorC[36] := BenchUut5.SensorC;
   TraceIn_ButtonA[36] := BenchUut5.ButtonA;
   TraceIn_ButtonB[36] := BenchUut5.ButtonB;
   TraceIn_ButtonC[36] := BenchUut5.ButtonC;
   BenchUut5();
   TraceOut_MotorForward[36] := BenchUut5.MotorForward;
   TraceOut_MotorReverse[36] := BenchUut5.MotorReverse;
   TraceOut_CompletionLight[36] := BenchUut5.CompletionLight;
   BenchCalls := BenchCalls + 1;
 37:
   BenchUut5.Mode := FALSE;
   BenchUut5.ForwardButton := TRUE;
   BenchUut5.ReverseButton := FALSE;
   BenchUut5.SensorA := FALSE;
   BenchUut5.SensorB := FALSE;
   BenchUut5.SensorC := FALSE;
   BenchUut5.ButtonA := FALSE;
   BenchUut5.ButtonB := FALSE;
   BenchUut5.ButtonC := FALSE;
   TraceIn_Mode[37] := BenchUut5.Mode;
   TraceIn_ForwardButton[37] := BenchUut5.ForwardButton;
   TraceIn_ReverseButton[37] := BenchUut5.ReverseButton;
   TraceIn_SensorA[37] := BenchUut5.SensorA;
   TraceIn_SensorB[37] := BenchUut5.SensorB;
   TraceIn_SensorC[37] := BenchUut5.SensorC;
   TraceIn_ButtonA[37] := BenchUut5.ButtonA;
   TraceIn_ButtonB[37] := BenchUut5.ButtonB;
   TraceIn_ButtonC[37] := BenchUut5.ButtonC;
   BenchUut5();
   TraceOut_MotorForward[37] := BenchUut5.MotorForward;
   TraceOut_MotorReverse[37] := BenchUut5.MotorReverse;
   TraceOut_CompletionLight[37] := BenchUut5.CompletionLight;
   BenchCalls := BenchCalls + 1;
 38:
   BenchUut5.Mode := FALSE;
   BenchUut5.ForwardButton := TRUE;
   BenchUut5.ReverseButton := FALSE;
   BenchUut5.SensorA := FALSE;
   BenchUut5.SensorB := FALSE;
   BenchUut5.SensorC := FALSE;
   BenchUut5.ButtonA := FALSE;
   BenchUut5.ButtonB := FALSE;
   BenchUut5.ButtonC := FALSE;
   TraceIn_Mode[38] := BenchUut5.Mode;
   TraceIn_ForwardButton[38] := BenchUut5.ForwardButton;
   TraceIn_ReverseButton[38] := BenchUut5.ReverseButton;
   TraceIn_SensorA[38] := BenchUut5.SensorA;
   TraceIn_SensorB[38] := BenchUut5.SensorB;
   TraceIn_SensorC[38] := BenchUut5.SensorC;
   TraceIn_ButtonA[38] := BenchUut5.ButtonA;
   TraceIn_ButtonB[38] := BenchUut5.ButtonB;
   TraceIn_ButtonC[38] := BenchUut5.ButtonC;
   BenchUut5();
   TraceOut_MotorForward[38] := BenchUut5.MotorForward;
   TraceOut_MotorReverse[38] := BenchUut5.MotorReverse;
   TraceOut_CompletionLight[38] := BenchUut5.CompletionLight;
   BenchCalls := BenchCalls + 1;
 39:
   BenchUut5.Mode := FALSE;
   BenchUut5.ForwardButton := TRUE;
   BenchUut5.ReverseButton := FALSE;
   BenchUut5.SensorA := FALSE;
   BenchUut5.SensorB := FALSE;
   BenchUut5.SensorC := FALSE;
   BenchUut5.ButtonA := FALSE;
   BenchUut5.ButtonB := FALSE;
   BenchUut5.ButtonC := FALSE;
   TraceIn_Mode[39] := BenchUut5.Mode;
   TraceIn_ForwardButton[39] := BenchUut5.ForwardButton;
   TraceIn_ReverseButton[39] := BenchUut5.ReverseButton;
   TraceIn_SensorA[39] := BenchUut5.SensorA;
   TraceIn_SensorB[39] := BenchUut5.SensorB;
   TraceIn_SensorC[39] := BenchUut5.SensorC;
   TraceIn_ButtonA[39] := BenchUut5.ButtonA;
   TraceIn_ButtonB[39] := BenchUut5.ButtonB;
   TraceIn_ButtonC[39] := BenchUut5.ButtonC;
   BenchUut5();
   TraceOut_MotorForward[39] := BenchUut5.MotorForward;
   TraceOut_MotorReverse[39] := BenchUut5.MotorReverse;
   TraceOut_CompletionLight[39] := BenchUut5.CompletionLight;
   BenchCalls := BenchCalls + 1;
 40:
   BenchUut5.Mode := FALSE;
   BenchUut5.ForwardButton := FALSE;
   BenchUut5.ReverseButton := TRUE;
   BenchUut5.SensorA := FALSE;
   BenchUut5.SensorB := FALSE;
   BenchUut5.SensorC := FALSE;
   BenchUut5.ButtonA := FALSE;
   BenchUut5.ButtonB := FALSE;
   BenchUut5.ButtonC := FALSE;
   TraceIn_Mode[40] := BenchUut5.Mode;
   TraceIn_ForwardButton[40] := BenchUut5.ForwardButton;
   TraceIn_ReverseButton[40] := BenchUut5.ReverseButton;
   TraceIn_SensorA[40] := BenchUut5.SensorA;
   TraceIn_SensorB[40] := BenchUut5.SensorB;
   TraceIn_SensorC[40] := BenchUut5.SensorC;
   TraceIn_ButtonA[40] := BenchUut5.ButtonA;
   TraceIn_ButtonB[40] := BenchUut5.ButtonB;
   TraceIn_ButtonC[40] := BenchUut5.ButtonC;
   BenchUut5();
   TraceOut_MotorForward[40] := BenchUut5.MotorForward;
   TraceOut_MotorReverse[40] := BenchUut5.MotorReverse;
   TraceOut_CompletionLight[40] := BenchUut5.CompletionLight;
   BenchCalls := BenchCalls + 1;
 41:
   BenchUut5.Mode := FALSE;
   BenchUut5.ForwardButton := FALSE;
   BenchUut5.ReverseButton := TRUE;
   BenchUut5.SensorA := FALSE;
   BenchUut5.SensorB := FALSE;
   BenchUut5.SensorC := FALSE;
   BenchUut5.ButtonA := FALSE;
   BenchUut5.ButtonB := FALSE;
   BenchUut5.ButtonC := FALSE;
   TraceIn_Mode[41] := BenchUut5.Mode;
   TraceIn_ForwardButton[41] := BenchUut5.ForwardButton;
   TraceIn_ReverseButton[41] := BenchUut5.ReverseButton;
   TraceIn_SensorA[41] := BenchUut5.SensorA;
   TraceIn_SensorB[41] := BenchUut5.SensorB;
   TraceIn_SensorC[41] := BenchUut5.SensorC;
   TraceIn_ButtonA[41] := BenchUut5.ButtonA;
   TraceIn_ButtonB[41] := BenchUut5.ButtonB;
   TraceIn_ButtonC[41] := BenchUut5.ButtonC;
   BenchUut5();
   TraceOut_MotorForward[41] := BenchUut5.MotorForward;
   TraceOut_MotorReverse[41] := BenchUut5.MotorReverse;
   TraceOut_CompletionLight[41] := BenchUut5.CompletionLight;
   BenchCalls := BenchCalls + 1;
 42:
   BenchUut5.Mode := FALSE;
   BenchUut5.ForwardButton := FALSE;
   BenchUut5.ReverseButton := TRUE;
   BenchUut5.SensorA := FALSE;
   BenchUut5.SensorB := FALSE;
   BenchUut5.SensorC := FALSE;
   BenchUut5.ButtonA := FALSE;
   BenchUut5.ButtonB := FALSE;
   BenchUut5.ButtonC := FALSE;
   TraceIn_Mode[42] := BenchUut5.Mode;
   TraceIn_ForwardButton[42] := BenchUut5.ForwardButton;
   TraceIn_ReverseButton[42] := BenchUut5.ReverseButton;
   TraceIn_SensorA[42] := BenchUut5.SensorA;
   TraceIn_SensorB[42] := BenchUut5.SensorB;
   TraceIn_SensorC[42] := BenchUut5.SensorC;
   TraceIn_ButtonA[42] := BenchUut5.ButtonA;
   TraceIn_ButtonB[42] := BenchUut5.ButtonB;
   TraceIn_ButtonC[42] := BenchUut5.ButtonC;
   BenchUut5();
   TraceOut_MotorForward[42] := BenchUut5.MotorForward;
   TraceOut_MotorReverse[42] := BenchUut5.MotorReverse;
   TraceOut_CompletionLight[42] := BenchUut5.CompletionLight;
   BenchCalls := BenchCalls + 1;
 43:
   BenchUut5.Mode := FALSE;
   BenchUut5.ForwardButton := TRUE;
   BenchUut5.ReverseButton := TRUE;
   BenchUut5.SensorA := FALSE;
   BenchUut5.SensorB := FALSE;
   BenchUut5.SensorC := FALSE;
   BenchUut5.ButtonA := FALSE;
   BenchUut5.ButtonB := FALSE;
   BenchUut5.ButtonC := FALSE;
   TraceIn_Mode[43] := BenchUut5.Mode;
   TraceIn_ForwardButton[43] := BenchUut5.ForwardButton;
   TraceIn_ReverseButton[43] := BenchUut5.ReverseButton;
   TraceIn_SensorA[43] := BenchUut5.SensorA;
   TraceIn_SensorB[43] := BenchUut5.SensorB;
   TraceIn_SensorC[43] := BenchUut5.SensorC;
   TraceIn_ButtonA[43] := BenchUut5.ButtonA;
   TraceIn_ButtonB[43] := BenchUut5.ButtonB;
   TraceIn_ButtonC[43] := BenchUut5.ButtonC;
   BenchUut5();
   TraceOut_MotorForward[43] := BenchUut5.MotorForward;
   TraceOut_MotorReverse[43] := BenchUut5.MotorReverse;
   TraceOut_CompletionLight[43] := BenchUut5.CompletionLight;
   BenchCalls := BenchCalls + 1;
 44:
   BenchUut5.Mode := FALSE;
   BenchUut5.ForwardButton := TRUE;
   BenchUut5.ReverseButton := TRUE;
   BenchUut5.SensorA := FALSE;
   BenchUut5.SensorB := FALSE;
   BenchUut5.SensorC := FALSE;
   BenchUut5.ButtonA := FALSE;
   BenchUut5.ButtonB := FALSE;
   BenchUut5.ButtonC := FALSE;
   TraceIn_Mode[44] := BenchUut5.Mode;
   TraceIn_ForwardButton[44] := BenchUut5.ForwardButton;
   TraceIn_ReverseButton[44] := BenchUut5.ReverseButton;
   TraceIn_SensorA[44] := BenchUut5.SensorA;
   TraceIn_SensorB[44] := BenchUut5.SensorB;
   TraceIn_SensorC[44] := BenchUut5.SensorC;
   TraceIn_ButtonA[44] := BenchUut5.ButtonA;
   TraceIn_ButtonB[44] := BenchUut5.ButtonB;
   TraceIn_ButtonC[44] := BenchUut5.ButtonC;
   BenchUut5();
   TraceOut_MotorForward[44] := BenchUut5.MotorForward;
   TraceOut_MotorReverse[44] := BenchUut5.MotorReverse;
   TraceOut_CompletionLight[44] := BenchUut5.CompletionLight;
   BenchCalls := BenchCalls + 1;
 45:
   BenchUut5.Mode := FALSE;
   BenchUut5.ForwardButton := TRUE;
   BenchUut5.ReverseButton := TRUE;
   BenchUut5.SensorA := FALSE;
   BenchUut5.SensorB := FALSE;
   BenchUut5.SensorC := FALSE;
   BenchUut5.ButtonA := FALSE;
   BenchUut5.ButtonB := FALSE;
   BenchUut5.ButtonC := FALSE;
   TraceIn_Mode[45] := BenchUut5.Mode;
   TraceIn_ForwardButton[45] := BenchUut5.ForwardButton;
   TraceIn_ReverseButton[45] := BenchUut5.ReverseButton;
   TraceIn_SensorA[45] := BenchUut5.SensorA;
   TraceIn_SensorB[45] := BenchUut5.SensorB;
   TraceIn_SensorC[45] := BenchUut5.SensorC;
   TraceIn_ButtonA[45] := BenchUut5.ButtonA;
   TraceIn_ButtonB[45] := BenchUut5.ButtonB;
   TraceIn_ButtonC[45] := BenchUut5.ButtonC;
   BenchUut5();
   TraceOut_MotorForward[45] := BenchUut5.MotorForward;
   TraceOut_MotorReverse[45] := BenchUut5.MotorReverse;
   TraceOut_CompletionLight[45] := BenchUut5.CompletionLight;
   BenchCalls := BenchCalls + 1;
 46:
   BenchUut6.Mode := TRUE;
   BenchUut6.ForwardButton := FALSE;
   BenchUut6.ReverseButton := FALSE;
   BenchUut6.SensorA := FALSE;
   BenchUut6.SensorB := FALSE;
   BenchUut6.SensorC := FALSE;
   BenchUut6.ButtonA := FALSE;
   BenchUut6.ButtonB := FALSE;
   BenchUut6.ButtonC := FALSE;
   TraceIn_Mode[46] := BenchUut6.Mode;
   TraceIn_ForwardButton[46] := BenchUut6.ForwardButton;
   TraceIn_ReverseButton[46] := BenchUut6.ReverseButton;
   TraceIn_SensorA[46] := BenchUut6.SensorA;
   TraceIn_SensorB[46] := BenchUut6.SensorB;
   TraceIn_SensorC[46] := BenchUut6.SensorC;
   TraceIn_ButtonA[46] := BenchUut6.ButtonA;
   TraceIn_ButtonB[46] := BenchUut6.ButtonB;
   TraceIn_ButtonC[46] := BenchUut6.ButtonC;
   BenchUut6();
   TraceOut_MotorForward[46] := BenchUut6.MotorForward;
   TraceOut_MotorReverse[46] := BenchUut6.MotorReverse;
   TraceOut_CompletionLight[46] := BenchUut6.CompletionLight;
   BenchCalls := BenchCalls + 1;
 47:
   BenchUut6.Mode := TRUE;
   BenchUut6.ForwardButton := FALSE;
   BenchUut6.ReverseButton := FALSE;
   BenchUut6.SensorA := FALSE;
   BenchUut6.SensorB := FALSE;
   BenchUut6.SensorC := FALSE;
   BenchUut6.ButtonA := FALSE;
   BenchUut6.ButtonB := FALSE;
   BenchUut6.ButtonC := FALSE;
   TraceIn_Mode[47] := BenchUut6.Mode;
   TraceIn_ForwardButton[47] := BenchUut6.ForwardButton;
   TraceIn_ReverseButton[47] := BenchUut6.ReverseButton;
   TraceIn_SensorA[47] := BenchUut6.SensorA;
   TraceIn_SensorB[47] := BenchUut6.SensorB;
   TraceIn_SensorC[47] := BenchUut6.SensorC;
   TraceIn_ButtonA[47] := BenchUut6.ButtonA;
   TraceIn_ButtonB[47] := BenchUut6.ButtonB;
   TraceIn_ButtonC[47] := BenchUut6.ButtonC;
   BenchUut6();
   TraceOut_MotorForward[47] := BenchUut6.MotorForward;
   TraceOut_MotorReverse[47] := BenchUut6.MotorReverse;
   TraceOut_CompletionLight[47] := BenchUut6.CompletionLight;
   BenchCalls := BenchCalls + 1;
 48:
   BenchUut6.Mode := TRUE;
   BenchUut6.ForwardButton := FALSE;
   BenchUut6.ReverseButton := FALSE;
   BenchUut6.SensorA := FALSE;
   BenchUut6.SensorB := FALSE;
   BenchUut6.SensorC := FALSE;
   BenchUut6.ButtonA := FALSE;
   BenchUut6.ButtonB := FALSE;
   BenchUut6.ButtonC := FALSE;
   TraceIn_Mode[48] := BenchUut6.Mode;
   TraceIn_ForwardButton[48] := BenchUut6.ForwardButton;
   TraceIn_ReverseButton[48] := BenchUut6.ReverseButton;
   TraceIn_SensorA[48] := BenchUut6.SensorA;
   TraceIn_SensorB[48] := BenchUut6.SensorB;
   TraceIn_SensorC[48] := BenchUut6.SensorC;
   TraceIn_ButtonA[48] := BenchUut6.ButtonA;
   TraceIn_ButtonB[48] := BenchUut6.ButtonB;
   TraceIn_ButtonC[48] := BenchUut6.ButtonC;
   BenchUut6();
   TraceOut_MotorForward[48] := BenchUut6.MotorForward;
   TraceOut_MotorReverse[48] := BenchUut6.MotorReverse;
   TraceOut_CompletionLight[48] := BenchUut6.CompletionLight;
   BenchCalls := BenchCalls + 1;
 49:
   BenchUut6.Mode := TRUE;
   BenchUut6.ForwardButton := FALSE;
   BenchUut6.ReverseButton := FALSE;
   BenchUut6.SensorA := TRUE;
   BenchUut6.SensorB := FALSE;
   BenchUut6.SensorC := FALSE;
   BenchUut6.ButtonA := FALSE;
   BenchUut6.ButtonB := FALSE;
   BenchUut6.ButtonC := FALSE;
   TraceIn_Mode[49] := BenchUut6.Mode;
   TraceIn_ForwardButton[49] := BenchUut6.ForwardButton;
   TraceIn_ReverseButton[49] := BenchUut6.ReverseButton;
   TraceIn_SensorA[49] := BenchUut6.SensorA;
   TraceIn_SensorB[49] := BenchUut6.SensorB;
   TraceIn_SensorC[49] := BenchUut6.SensorC;
   TraceIn_ButtonA[49] := BenchUut6.ButtonA;
   TraceIn_ButtonB[49] := BenchUut6.ButtonB;
   TraceIn_ButtonC[49] := BenchUut6.ButtonC;
   BenchUut6();
   TraceOut_MotorForward[49] := BenchUut6.MotorForward;
   TraceOut_MotorReverse[49] := BenchUut6.MotorReverse;
   TraceOut_CompletionLight[49] := BenchUut6.CompletionLight;
   BenchCalls := BenchCalls + 1;
 50:
   BenchUut6.Mode := TRUE;
   BenchUut6.ForwardButton := FALSE;
   BenchUut6.ReverseButton := FALSE;
   BenchUut6.SensorA := TRUE;
   BenchUut6.SensorB := FALSE;
   BenchUut6.SensorC := FALSE;
   BenchUut6.ButtonA := FALSE;
   BenchUut6.ButtonB := FALSE;
   BenchUut6.ButtonC := FALSE;
   TraceIn_Mode[50] := BenchUut6.Mode;
   TraceIn_ForwardButton[50] := BenchUut6.ForwardButton;
   TraceIn_ReverseButton[50] := BenchUut6.ReverseButton;
   TraceIn_SensorA[50] := BenchUut6.SensorA;
   TraceIn_SensorB[50] := BenchUut6.SensorB;
   TraceIn_SensorC[50] := BenchUut6.SensorC;
   TraceIn_ButtonA[50] := BenchUut6.ButtonA;
   TraceIn_ButtonB[50] := BenchUut6.ButtonB;
   TraceIn_ButtonC[50] := BenchUut6.ButtonC;
   BenchUut6();
   TraceOut_MotorForward[50] := BenchUut6.MotorForward;
   TraceOut_MotorReverse[50] := BenchUut6.MotorReverse;
   TraceOut_CompletionLight[50] := BenchUut6.CompletionLight;
   BenchCalls := BenchCalls + 1;
 51:
   BenchUut6.Mode := TRUE;
   BenchUut6.ForwardButton := FALSE;
   BenchUut6.ReverseButton := FALSE;
   BenchUut6.SensorA := TRUE;
   BenchUut6.SensorB := FALSE;
   BenchUut6.SensorC := FALSE;
   BenchUut6.ButtonA := FALSE;
   BenchUut6.ButtonB := FALSE;
   BenchUut6.ButtonC := FALSE;
   TraceIn_Mode[51] := BenchUut6.Mode;
   TraceIn_ForwardButton[51] := BenchUut6.ForwardButton;
   TraceIn_ReverseButton[51] := BenchUut6.ReverseButton;
   TraceIn_SensorA[51] := BenchUut6.SensorA;
   TraceIn_SensorB[51] := BenchUut6.SensorB;
   TraceIn_SensorC[51] := BenchUut6.SensorC;
   TraceIn_ButtonA[51] := BenchUut6.ButtonA;
   TraceIn_ButtonB[51] := BenchUut6.ButtonB;
   TraceIn_ButtonC[51] := BenchUut6.ButtonC;
   BenchUut6();
   TraceOut_MotorForward[51] := BenchUut6.MotorForward;
   TraceOut_MotorReverse[51] := BenchUut6.MotorReverse;
   TraceOut_CompletionLight[51] := BenchUut6.CompletionLight;
   BenchCalls := BenchCalls + 1;
 52:
   BenchUut6.Mode := TRUE;
   BenchUut6.ForwardButton := FALSE;
   BenchUut6.ReverseButton := FALSE;
   BenchUut6.SensorA := TRUE;
   BenchUut6.SensorB := FALSE;
   BenchUut6.SensorC := FALSE;
   BenchUut6.ButtonA := TRUE;
   BenchUut6.ButtonB := FALSE;
   BenchUut6.ButtonC := FALSE;
   TraceIn_Mode[52] := BenchUut6.Mode;
   TraceIn_ForwardButton[52] := BenchUut6.ForwardButton;
   TraceIn_ReverseButton[52] := BenchUut6.ReverseButton;
   TraceIn_SensorA[52] := BenchUut6.SensorA;
   TraceIn_SensorB[52] := BenchUut6.SensorB;
   TraceIn_SensorC[52] := BenchUut6.SensorC;
   TraceIn_ButtonA[52] := BenchUut6.ButtonA;
   TraceIn_ButtonB[52] := BenchUut6.ButtonB;
   TraceIn_ButtonC[52] := BenchUut6.ButtonC;
   BenchUut6();
   TraceOut_MotorForward[52] := BenchUut6.MotorForward;
   TraceOut_MotorReverse[52] := BenchUut6.MotorReverse;
   TraceOut_CompletionLight[52] := BenchUut6.CompletionLight;
   BenchCalls := BenchCalls + 1;
 53:
   BenchUut6.Mode := TRUE;
   BenchUut6.ForwardButton := FALSE;
   BenchUut6.ReverseButton := FALSE;
   BenchUut6.SensorA := TRUE;
   BenchUut6.SensorB := FALSE;
   BenchUut6.SensorC := FALSE;
   BenchUut6.ButtonA := TRUE;
   BenchUut6.ButtonB := FALSE;
   BenchUut6.ButtonC := FALSE;
   TraceIn_Mode[53] := BenchUut6.Mode;
   TraceIn_ForwardButton[53] := BenchUut6.ForwardButton;
   TraceIn_ReverseButton[53] := BenchUut6.ReverseButton;
   TraceIn_SensorA[53] := BenchUut6.SensorA;
   TraceIn_SensorB[53] := BenchUut6.SensorB;
   TraceIn_SensorC[53] := BenchUut6.SensorC;
   TraceIn_ButtonA[53] := BenchUut6.ButtonA;
   TraceIn_ButtonB[53] := BenchUut6.ButtonB;
   TraceIn_ButtonC[53] := BenchUut6.ButtonC;
   BenchUut6();
   TraceOut_MotorForward[53] := BenchUut6.MotorForward;
   TraceOut_MotorReverse[53] := BenchUut6.MotorReverse;
   TraceOut_CompletionLight[53] := BenchUut6.CompletionLight;
   BenchCalls := BenchCalls + 1;
 54:
   BenchUut6.Mode := TRUE;
   BenchUut6.ForwardButton := FALSE;
   BenchUut6.ReverseButton := FALSE;
   BenchUut6.SensorA := TRUE;
   BenchUut6.SensorB := FALSE;
   BenchUut6.SensorC := FALSE;
   BenchUut6.ButtonA := TRUE;
   BenchUut6.ButtonB := FALSE;
   BenchUut6.ButtonC := FALSE;
   TraceIn_Mode[54] := BenchUut6.Mode;
   TraceIn_ForwardButton[54] := BenchUut6.ForwardButton;
   TraceIn_ReverseButton[54] := BenchUut6.ReverseButton;
   TraceIn_SensorA[54] := BenchUut6.SensorA;
   TraceIn_SensorB[54] := BenchUut6.SensorB;
   TraceIn_SensorC[54] := BenchUut6.SensorC;
   TraceIn_ButtonA[54] := BenchUut6.ButtonA;
   TraceIn_ButtonB[54] := BenchUut6.ButtonB;
   TraceIn_ButtonC[54] := BenchUut6.ButtonC;
   BenchUut6();
   TraceOut_MotorForward[54] := BenchUut6.MotorForward;
   TraceOut_MotorReverse[54] := BenchUut6.MotorReverse;
   TraceOut_CompletionLight[54] := BenchUut6.CompletionLight;
   BenchCalls := BenchCalls + 1;
 55:
   BenchUut6.Mode := TRUE;
   BenchUut6.ForwardButton := FALSE;
   BenchUut6.ReverseButton := FALSE;
   BenchUut6.SensorA := FALSE;
   BenchUut6.SensorB := FALSE;
   BenchUut6.SensorC := FALSE;
   BenchUut6.ButtonA := FALSE;
   BenchUut6.ButtonB := FALSE;
   BenchUut6.ButtonC := FALSE;
   TraceIn_Mode[55] := BenchUut6.Mode;
   TraceIn_ForwardButton[55] := BenchUut6.ForwardButton;
   TraceIn_ReverseButton[55] := BenchUut6.ReverseButton;
   TraceIn_SensorA[55] := BenchUut6.SensorA;
   TraceIn_SensorB[55] := BenchUut6.SensorB;
   TraceIn_SensorC[55] := BenchUut6.SensorC;
   TraceIn_ButtonA[55] := BenchUut6.ButtonA;
   TraceIn_ButtonB[55] := BenchUut6.ButtonB;
   TraceIn_ButtonC[55] := BenchUut6.ButtonC;
   BenchUut6();
   TraceOut_MotorForward[55] := BenchUut6.MotorForward;
   TraceOut_MotorReverse[55] := BenchUut6.MotorReverse;
   TraceOut_CompletionLight[55] := BenchUut6.CompletionLight;
   BenchCalls := BenchCalls + 1;
 56:
   BenchUut6.Mode := TRUE;
   BenchUut6.ForwardButton := FALSE;
   BenchUut6.ReverseButton := FALSE;
   BenchUut6.SensorA := FALSE;
   BenchUut6.SensorB := FALSE;
   BenchUut6.SensorC := FALSE;
   BenchUut6.ButtonA := FALSE;
   BenchUut6.ButtonB := FALSE;
   BenchUut6.ButtonC := FALSE;
   TraceIn_Mode[56] := BenchUut6.Mode;
   TraceIn_ForwardButton[56] := BenchUut6.ForwardButton;
   TraceIn_ReverseButton[56] := BenchUut6.ReverseButton;
   TraceIn_SensorA[56] := BenchUut6.SensorA;
   TraceIn_SensorB[56] := BenchUut6.SensorB;
   TraceIn_SensorC[56] := BenchUut6.SensorC;
   TraceIn_ButtonA[56] := BenchUut6.ButtonA;
   TraceIn_ButtonB[56] := BenchUut6.ButtonB;
   TraceIn_ButtonC[56] := BenchUut6.ButtonC;
   BenchUut6();
   TraceOut_MotorForward[56] := BenchUut6.MotorForward;
   TraceOut_MotorReverse[56] := BenchUut6.MotorReverse;
   TraceOut_CompletionLight[56] := BenchUut6.CompletionLight;
   BenchCalls := BenchCalls + 1;
 57:
   BenchUut6.Mode := TRUE;
   BenchUut6.ForwardButton := FALSE;
   BenchUut6.ReverseButton := FALSE;
   BenchUut6.SensorA := FALSE;
   BenchUut6.SensorB := FALSE;
   BenchUut6.SensorC := FALSE;
   BenchUut6.ButtonA := FALSE;
   BenchUut6.ButtonB := FALSE;
   BenchUut6.ButtonC := FALSE;
   TraceIn_Mode[57] := BenchUut6.Mode;
   TraceIn_ForwardButton[57] := BenchUut6.ForwardButton;
   TraceIn_ReverseButton[57] := BenchUut6.ReverseButton;
   TraceIn_SensorA[57] := BenchUut6.SensorA;
   TraceIn_SensorB[57] := BenchUut6.SensorB;
   TraceIn_SensorC[57] := BenchUut6.SensorC;
   TraceIn_ButtonA[57] := BenchUut6.ButtonA;
   TraceIn_ButtonB[57] := BenchUut6.ButtonB;
   TraceIn_ButtonC[57] := BenchUut6.ButtonC;
   BenchUut6();
   TraceOut_MotorForward[57] := BenchUut6.MotorForward;
   TraceOut_MotorReverse[57] := BenchUut6.MotorReverse;
   TraceOut_CompletionLight[57] := BenchUut6.CompletionLight;
   BenchCalls := BenchCalls + 1;
 58:
   BenchUut6.Mode := TRUE;
   BenchUut6.ForwardButton := FALSE;
   BenchUut6.ReverseButton := FALSE;
   BenchUut6.SensorA := FALSE;
   BenchUut6.SensorB := TRUE;
   BenchUut6.SensorC := FALSE;
   BenchUut6.ButtonA := FALSE;
   BenchUut6.ButtonB := FALSE;
   BenchUut6.ButtonC := FALSE;
   TraceIn_Mode[58] := BenchUut6.Mode;
   TraceIn_ForwardButton[58] := BenchUut6.ForwardButton;
   TraceIn_ReverseButton[58] := BenchUut6.ReverseButton;
   TraceIn_SensorA[58] := BenchUut6.SensorA;
   TraceIn_SensorB[58] := BenchUut6.SensorB;
   TraceIn_SensorC[58] := BenchUut6.SensorC;
   TraceIn_ButtonA[58] := BenchUut6.ButtonA;
   TraceIn_ButtonB[58] := BenchUut6.ButtonB;
   TraceIn_ButtonC[58] := BenchUut6.ButtonC;
   BenchUut6();
   TraceOut_MotorForward[58] := BenchUut6.MotorForward;
   TraceOut_MotorReverse[58] := BenchUut6.MotorReverse;
   TraceOut_CompletionLight[58] := BenchUut6.CompletionLight;
   BenchCalls := BenchCalls + 1;
 59:
   BenchUut6.Mode := TRUE;
   BenchUut6.ForwardButton := FALSE;
   BenchUut6.ReverseButton := FALSE;
   BenchUut6.SensorA := FALSE;
   BenchUut6.SensorB := TRUE;
   BenchUut6.SensorC := FALSE;
   BenchUut6.ButtonA := FALSE;
   BenchUut6.ButtonB := FALSE;
   BenchUut6.ButtonC := FALSE;
   TraceIn_Mode[59] := BenchUut6.Mode;
   TraceIn_ForwardButton[59] := BenchUut6.ForwardButton;
   TraceIn_ReverseButton[59] := BenchUut6.ReverseButton;
   TraceIn_SensorA[59] := BenchUut6.SensorA;
   TraceIn_SensorB[59] := BenchUut6.SensorB;
   TraceIn_SensorC[59] := BenchUut6.SensorC;
   TraceIn_ButtonA[59] := BenchUut6.ButtonA;
   TraceIn_ButtonB[59] := BenchUut6.ButtonB;
   TraceIn_ButtonC[59] := BenchUut6.ButtonC;
   BenchUut6();
   TraceOut_MotorForward[59] := BenchUut6.MotorForward;
   TraceOut_MotorReverse[59] := BenchUut6.MotorReverse;
   TraceOut_CompletionLight[59] := BenchUut6.CompletionLight;
   BenchCalls := BenchCalls + 1;
 60:
   BenchUut6.Mode := TRUE;
   BenchUut6.ForwardButton := FALSE;
   BenchUut6.ReverseButton := FALSE;
   BenchUut6.SensorA := FALSE;
   BenchUut6.SensorB := TRUE;
   BenchUut6.SensorC := FALSE;
   BenchUut6.ButtonA := FALSE;
   BenchUut6.ButtonB := FALSE;
   BenchUut6.ButtonC := FALSE;
   TraceIn_Mode[60] := BenchUut6.Mode;
   TraceIn_ForwardButton[60] := BenchUut6.ForwardButton;
   TraceIn_ReverseButton[60] := BenchUut6.ReverseButton;
   TraceIn_SensorA[60] := BenchUut6.SensorA;
   TraceIn_SensorB[60] := BenchUut6.SensorB;
   TraceIn_SensorC[60] := BenchUut6.SensorC;
   TraceIn_ButtonA[60] := BenchUut6.ButtonA;
   TraceIn_ButtonB[60] := BenchUut6.ButtonB;
   TraceIn_ButtonC[60] := BenchUut6.ButtonC;
   BenchUut6();
   TraceOut_MotorForward[60] := BenchUut6.MotorForward;
   TraceOut_MotorReverse[60] := BenchUut6.MotorReverse;
   TraceOut_CompletionLight[60] := BenchUut6.CompletionLight;
   BenchCalls := BenchCalls + 1;
 61:
   BenchUut6.Mode := TRUE;
   BenchUut6.ForwardButton := FALSE;
   BenchUut6.ReverseButton := FALSE;
   BenchUut6.SensorA := FALSE;
   BenchUut6.SensorB := TRUE;
   BenchUut6.SensorC := FALSE;
   BenchUut6.ButtonA := FALSE;
   BenchUut6.ButtonB := TRUE;
   BenchUut6.ButtonC := FALSE;
   TraceIn_Mode[61] := BenchUut6.Mode;
   TraceIn_ForwardButton[61] := BenchUut6.ForwardButton;
   TraceIn_ReverseButton[61] := BenchUut6.ReverseButton;
   TraceIn_SensorA[61] := BenchUut6.SensorA;
   TraceIn_SensorB[61] := BenchUut6.SensorB;
   TraceIn_SensorC[61] := BenchUut6.SensorC;
   TraceIn_ButtonA[61] := BenchUut6.ButtonA;
   TraceIn_ButtonB[61] := BenchUut6.ButtonB;
   TraceIn_ButtonC[61] := BenchUut6.ButtonC;
   BenchUut6();
   TraceOut_MotorForward[61] := BenchUut6.MotorForward;
   TraceOut_MotorReverse[61] := BenchUut6.MotorReverse;
   TraceOut_CompletionLight[61] := BenchUut6.CompletionLight;
   BenchCalls := BenchCalls + 1;
 62:
   BenchUut6.Mode := TRUE;
   BenchUut6.ForwardButton := FALSE;
   BenchUut6.ReverseButton := FALSE;
   BenchUut6.SensorA := FALSE;
   BenchUut6.SensorB := TRUE;
   BenchUut6.SensorC := FALSE;
   BenchUut6.ButtonA := FALSE;
   BenchUut6.ButtonB := TRUE;
   BenchUut6.ButtonC := FALSE;
   TraceIn_Mode[62] := BenchUut6.Mode;
   TraceIn_ForwardButton[62] := BenchUut6.ForwardButton;
   TraceIn_ReverseButton[62] := BenchUut6.ReverseButton;
   TraceIn_SensorA[62] := BenchUut6.SensorA;
   TraceIn_SensorB[62] := BenchUut6.SensorB;
   TraceIn_SensorC[62] := BenchUut6.SensorC;
   TraceIn_ButtonA[62] := BenchUut6.ButtonA;
   TraceIn_ButtonB[62] := BenchUut6.ButtonB;
   TraceIn_ButtonC[62] := BenchUut6.ButtonC;
   BenchUut6();
   TraceOut_MotorForward[62] := BenchUut6.MotorForward;
   TraceOut_MotorReverse[62] := BenchUut6.MotorReverse;
   TraceOut_CompletionLight[62] := BenchUut6.CompletionLight;
   BenchCalls := BenchCalls + 1;
 63:
   BenchUut6.Mode := TRUE;
   BenchUut6.ForwardButton := FALSE;
   BenchUut6.ReverseButton := FALSE;
   BenchUut6.SensorA := FALSE;
   BenchUut6.SensorB := TRUE;
   BenchUut6.SensorC := FALSE;
   BenchUut6.ButtonA := FALSE;
   BenchUut6.ButtonB := TRUE;
   BenchUut6.ButtonC := FALSE;
   TraceIn_Mode[63] := BenchUut6.Mode;
   TraceIn_ForwardButton[63] := BenchUut6.ForwardButton;
   TraceIn_ReverseButton[63] := BenchUut6.ReverseButton;
   TraceIn_SensorA[63] := BenchUut6.SensorA;
   TraceIn_SensorB[63] := BenchUut6.SensorB;
   TraceIn_SensorC[63] := BenchUut6.SensorC;
   TraceIn_ButtonA[63] := BenchUut6.ButtonA;
   TraceIn_ButtonB[63] := BenchUut6.ButtonB;
   TraceIn_ButtonC[63] := BenchUut6.ButtonC;
   BenchUut6();
   TraceOut_MotorForward[63] := BenchUut6.MotorForward;
   TraceOut_MotorReverse[63] := BenchUut6.MotorReverse;
   TraceOut_CompletionLight[63] := BenchUut6.CompletionLight;
   BenchCalls := BenchCalls + 1;
 64:
   BenchUut6.Mode := TRUE;
   BenchUut6.ForwardButton := FALSE;
   BenchUut6.ReverseButton := FALSE;
   BenchUut6.SensorA := FALSE;
   BenchUut6.SensorB := FALSE;
   BenchUut6.SensorC := TRUE;
   BenchUut6.ButtonA := FALSE;
   BenchUut6.ButtonB := FALSE;
   BenchUut6.ButtonC := FALSE;
   TraceIn_Mode[64] := BenchUut6.Mode;
   TraceIn_ForwardButton[64] := BenchUut6.ForwardButton;
   TraceIn_ReverseButton[64] := BenchUut6.ReverseButton;
   TraceIn_SensorA[64] := BenchUut6.SensorA;
   TraceIn_SensorB[64] := BenchUut6.SensorB;
   TraceIn_SensorC[64] := BenchUut6.SensorC;
   TraceIn_ButtonA[64] := BenchUut6.ButtonA;
   TraceIn_ButtonB[64] := BenchUut6.ButtonB;
   TraceIn_ButtonC[64] := BenchUut6.ButtonC;
   BenchUut6();
   TraceOut_MotorForward[64] := BenchUut6.MotorForward;
   TraceOut_MotorReverse[64] := BenchUut6.MotorReverse;
   TraceOut_CompletionLight[64] := BenchUut6.CompletionLight;
   BenchCalls := BenchCalls + 1;
 65:
   BenchUut6.Mode := TRUE;
   BenchUut6.ForwardButton := FALSE;
   BenchUut6.ReverseButton := FALSE;
   BenchUut6.SensorA := FALSE;
   BenchUut6.SensorB := FALSE;
   BenchUut6.SensorC := TRUE;
   BenchUut6.ButtonA := FALSE;
   BenchUut6.ButtonB := FALSE;
   BenchUut6.ButtonC := FALSE;
   TraceIn_Mode[65] := BenchUut6.Mode;
   TraceIn_ForwardButton[65] := BenchUut6.ForwardButton;
   TraceIn_ReverseButton[65] := BenchUut6.ReverseButton;
   TraceIn_SensorA[65] := BenchUut6.SensorA;
   TraceIn_SensorB[65] := BenchUut6.SensorB;
   TraceIn_SensorC[65] := BenchUut6.SensorC;
   TraceIn_ButtonA[65] := BenchUut6.ButtonA;
   TraceIn_ButtonB[65] := BenchUut6.ButtonB;
   TraceIn_ButtonC[65] := BenchUut6.ButtonC;
   BenchUut6();
   TraceOut_MotorForward[65] := BenchUut6.MotorForward;
   TraceOut_MotorReverse[65] := BenchUut6.MotorReverse;
   TraceOut_CompletionLight[65] := BenchUut6.CompletionLight;
   BenchCalls := BenchCalls + 1;
 66:
   BenchUut6.Mode := TRUE;
   BenchUut6.ForwardButton := FALSE;
   BenchUut6.ReverseButton := FALSE;
   BenchUut6.SensorA := FALSE;
   BenchUut6.SensorB := FALSE;
   BenchUut6.SensorC := TRUE;
   BenchUut6.ButtonA := FALSE;
   BenchUut6.ButtonB := FALSE;
   BenchUut6.ButtonC := FALSE;
   TraceIn_Mode[66] := BenchUut6.Mode;
   TraceIn_ForwardButton[66] := BenchUut6.ForwardButton;
   TraceIn_ReverseButton[66] := BenchUut6.ReverseButton;
   TraceIn_SensorA[66] := BenchUut6.SensorA;
   TraceIn_SensorB[66] := BenchUut6.SensorB;
   TraceIn_SensorC[66] := BenchUut6.SensorC;
   TraceIn_ButtonA[66] := BenchUut6.ButtonA;
   TraceIn_ButtonB[66] := BenchUut6.ButtonB;
   TraceIn_ButtonC[66] := BenchUut6.ButtonC;
   BenchUut6();
   TraceOut_MotorForward[66] := BenchUut6.MotorForward;
   TraceOut_MotorReverse[66] := BenchUut6.MotorReverse;
   TraceOut_CompletionLight[66] := BenchUut6.CompletionLight;
   BenchCalls := BenchCalls + 1;
 67:
   BenchUut6.Mode := TRUE;
   BenchUut6.ForwardButton := FALSE;
   BenchUut6.ReverseButton := FALSE;
   BenchUut6.SensorA := FALSE;
   BenchUut6.SensorB := FALSE;
   BenchUut6.SensorC := TRUE;
   BenchUut6.ButtonA := FALSE;
   BenchUut6.ButtonB := FALSE;
   BenchUut6.ButtonC := TRUE;
   TraceIn_Mode[67] := BenchUut6.Mode;
   TraceIn_ForwardButton[67] := BenchUut6.ForwardButton;
   TraceIn_ReverseButton[67] := BenchUut6.ReverseButton;
   TraceIn_SensorA[67] := BenchUut6.SensorA;
   TraceIn_SensorB[67] := BenchUut6.SensorB;
   TraceIn_SensorC[67] := BenchUut6.SensorC;
   TraceIn_ButtonA[67] := BenchUut6.ButtonA;
   TraceIn_ButtonB[67] := BenchUut6.ButtonB;
   TraceIn_ButtonC[67] := BenchUut6.ButtonC;
   BenchUut6();
   TraceOut_MotorForward[67] := BenchUut6.MotorForward;
   TraceOut_MotorReverse[67] := BenchUut6.MotorReverse;
   TraceOut_CompletionLight[67] := BenchUut6.CompletionLight;
   BenchCalls := BenchCalls + 1;
 68:
   BenchUut6.Mode := TRUE;
   BenchUut6.ForwardButton := FALSE;
   BenchUut6.ReverseButton := FALSE;
   BenchUut6.SensorA := FALSE;
   BenchUut6.SensorB := FALSE;
   BenchUut6.SensorC := TRUE;
   BenchUut6.ButtonA := FALSE;
   BenchUut6.ButtonB := FALSE;
   BenchUut6.ButtonC := TRUE;
   TraceIn_Mode[68] := BenchUut6.Mode;
   TraceIn_ForwardButton[68] := BenchUut6.ForwardButton;
   TraceIn_ReverseButton[68] := BenchUut6.ReverseButton;
   TraceIn_SensorA[68] := BenchUut6.SensorA;
   TraceIn_SensorB[68] := BenchUut6.SensorB;
   TraceIn_SensorC[68] := BenchUut6.SensorC;
   TraceIn_ButtonA[68] := BenchUut6.ButtonA;
   TraceIn_ButtonB[68] := BenchUut6.ButtonB;
   TraceIn_ButtonC[68] := BenchUut6.ButtonC;
   BenchUut6();
   TraceOut_MotorForward[68] := BenchUut6.MotorForward;
   TraceOut_MotorReverse[68] := BenchUut6.MotorReverse;
   TraceOut_CompletionLight[68] := BenchUut6.CompletionLight;
   BenchCalls := BenchCalls + 1;
 69:
   BenchUut6.Mode := TRUE;
   BenchUut6.ForwardButton := FALSE;
   BenchUut6.ReverseButton := FALSE;
   BenchUut6.SensorA := FALSE;
   BenchUut6.SensorB := FALSE;
   BenchUut6.SensorC := TRUE;
   BenchUut6.ButtonA := FALSE;
   BenchUut6.ButtonB := FALSE;
   BenchUut6.ButtonC := TRUE;
   TraceIn_Mode[69] := BenchUut6.Mode;
   TraceIn_ForwardButton[69] := BenchUut6.ForwardButton;
   TraceIn_ReverseButton[69] := BenchUut6.ReverseButton;
   TraceIn_SensorA[69] := BenchUut6.SensorA;
   TraceIn_SensorB[69] := BenchUut6.SensorB;
   TraceIn_SensorC[69] := BenchUut6.SensorC;
   TraceIn_ButtonA[69] := BenchUut6.ButtonA;
   TraceIn_ButtonB[69] := BenchUut6.ButtonB;
   TraceIn_ButtonC[69] := BenchUut6.ButtonC;
   BenchUut6();
   TraceOut_MotorForward[69] := BenchUut6.MotorForward;
   TraceOut_MotorReverse[69] := BenchUut6.MotorReverse;
   TraceOut_CompletionLight[69] := BenchUut6.CompletionLight;
   BenchCalls := BenchCalls + 1;
 70:
   BenchUut6.Mode := TRUE;
   BenchUut6.ForwardButton := FALSE;
   BenchUut6.ReverseButton := FALSE;
   BenchUut6.SensorA := FALSE;
   BenchUut6.SensorB := FALSE;
   BenchUut6.SensorC := TRUE;
   BenchUut6.ButtonA := FALSE;
   BenchUut6.ButtonB := FALSE;
   BenchUut6.ButtonC := FALSE;
   TraceIn_Mode[70] := BenchUut6.Mode;
   TraceIn_ForwardButton[70] := BenchUut6.ForwardButton;
   TraceIn_ReverseButton[70] := BenchUut6.ReverseButton;
   TraceIn_SensorA[70] := BenchUut6.SensorA;
   TraceIn_SensorB[70] := BenchUut6.SensorB;
   TraceIn_SensorC[70] := BenchUut6.SensorC;
   TraceIn_ButtonA[70] := BenchUut6.ButtonA;
   TraceIn_ButtonB[70] := BenchUut6.ButtonB;
   TraceIn_ButtonC[70] := BenchUut6.ButtonC;
   BenchUut6();
   TraceOut_MotorForward[70] := BenchUut6.MotorForward;
   TraceOut_MotorReverse[70] := BenchUut6.MotorReverse;
   TraceOut_CompletionLight[70] := BenchUut6.CompletionLight;
   BenchCalls := BenchCalls + 1;
 71:
   BenchUut6.Mode := TRUE;
   BenchUut6.ForwardButton := FALSE;
   BenchUut6.ReverseButton := FALSE;
   BenchUut6.SensorA := FALSE;
   BenchUut6.SensorB := FALSE;
   BenchUut6.SensorC := TRUE;
   BenchUut6.ButtonA := FALSE;
   BenchUut6.ButtonB := FALSE;
   BenchUut6.ButtonC := FALSE;
   TraceIn_Mode[71] := BenchUut6.Mode;
   TraceIn_ForwardButton[71] := BenchUut6.ForwardButton;
   TraceIn_ReverseButton[71] := BenchUut6.ReverseButton;
   TraceIn_SensorA[71] := BenchUut6.SensorA;
   TraceIn_SensorB[71] := BenchUut6.SensorB;
   TraceIn_SensorC[71] := BenchUut6.SensorC;
   TraceIn_ButtonA[71] := BenchUut6.ButtonA;
   TraceIn_ButtonB[71] := BenchUut6.ButtonB;
   TraceIn_ButtonC[71] := BenchUut6.ButtonC;
   BenchUut6();
   TraceOut_MotorForward[71] := BenchUut6.MotorForward;
   TraceOut_MotorReverse[71] := BenchUut6.MotorReverse;
   TraceOut_CompletionLight[71] := BenchUut6.CompletionLight;
   BenchCalls := BenchCalls + 1;
 72:
   BenchUut6.Mode := TRUE;
   BenchUut6.ForwardButton := FALSE;
   BenchUut6.ReverseButton := FALSE;
   BenchUut6.SensorA := FALSE;
   BenchUut6.SensorB := FALSE;
   BenchUut6.SensorC := TRUE;
   BenchUut6.ButtonA := FALSE;
   BenchUut6.ButtonB := FALSE;
   BenchUut6.ButtonC := FALSE;
   TraceIn_Mode[72] := BenchUut6.Mode;
   TraceIn_ForwardButton[72] := BenchUut6.ForwardButton;
   TraceIn_ReverseButton[72] := BenchUut6.ReverseButton;
   TraceIn_SensorA[72] := BenchUut6.SensorA;
   TraceIn_SensorB[72] := BenchUut6.SensorB;
   TraceIn_SensorC[72] := BenchUut6.SensorC;
   TraceIn_ButtonA[72] := BenchUut6.ButtonA;
   TraceIn_ButtonB[72] := BenchUut6.ButtonB;
   TraceIn_ButtonC[72] := BenchUut6.ButtonC;
   BenchUut6();
   TraceOut_MotorForward[72] := BenchUut6.MotorForward;
   TraceOut_MotorReverse[72] := BenchUut6.MotorReverse;
   TraceOut_CompletionLight[72] := BenchUut6.CompletionLight;
   BenchCalls := BenchCalls + 1;
 73:
   BenchUut6.Mode := TRUE;
   BenchUut6.ForwardButton := FALSE;
   BenchUut6.ReverseButton := FALSE;
   BenchUut6.SensorA := FALSE;
   BenchUut6.SensorB := FALSE;
   BenchUut6.SensorC := FALSE;
   BenchUut6.ButtonA := FALSE;
   BenchUut6.ButtonB := FALSE;
   BenchUut6.ButtonC := FALSE;
   TraceIn_Mode[73] := BenchUut6.Mode;
   TraceIn_ForwardButton[73] := BenchUut6.ForwardButton;
   TraceIn_ReverseButton[73] := BenchUut6.ReverseButton;
   TraceIn_SensorA[73] := BenchUut6.SensorA;
   TraceIn_SensorB[73] := BenchUut6.SensorB;
   TraceIn_SensorC[73] := BenchUut6.SensorC;
   TraceIn_ButtonA[73] := BenchUut6.ButtonA;
   TraceIn_ButtonB[73] := BenchUut6.ButtonB;
   TraceIn_ButtonC[73] := BenchUut6.ButtonC;
   BenchUut6();
   TraceOut_MotorForward[73] := BenchUut6.MotorForward;
   TraceOut_MotorReverse[73] := BenchUut6.MotorReverse;
   TraceOut_CompletionLight[73] := BenchUut6.CompletionLight;
   BenchCalls := BenchCalls + 1;
 74:
   BenchUut6.Mode := TRUE;
   BenchUut6.ForwardButton := FALSE;
   BenchUut6.ReverseButton := FALSE;
   BenchUut6.SensorA := FALSE;
   BenchUut6.SensorB := FALSE;
   BenchUut6.SensorC := FALSE;
   BenchUut6.ButtonA := FALSE;
   BenchUut6.ButtonB := FALSE;
   BenchUut6.ButtonC := FALSE;
   TraceIn_Mode[74] := BenchUut6.Mode;
   TraceIn_ForwardButton[74] := BenchUut6.ForwardButton;
   TraceIn_ReverseButton[74] := BenchUut6.ReverseButton;
   TraceIn_SensorA[74] := BenchUut6.SensorA;
   TraceIn_SensorB[74] := BenchUut6.SensorB;
   TraceIn_SensorC[74] := BenchUut6.SensorC;
   TraceIn_ButtonA[74] := BenchUut6.ButtonA;
   TraceIn_ButtonB[74] := BenchUut6.ButtonB;
   TraceIn_ButtonC[74] := BenchUut6.ButtonC;
   BenchUut6();
   TraceOut_MotorForward[74] := BenchUut6.MotorForward;
   TraceOut_MotorReverse[74] := BenchUut6.MotorReverse;
   TraceOut_CompletionLight[74] := BenchUut6.CompletionLight;
   BenchCalls := BenchCalls + 1;
 75:
   BenchUut6.Mode := TRUE;
   BenchUut6.ForwardButton := FALSE;
   BenchUut6.ReverseButton := FALSE;
   BenchUut6.SensorA := FALSE;
   BenchUut6.SensorB := FALSE;
   BenchUut6.SensorC := FALSE;
   BenchUut6.ButtonA := FALSE;
   BenchUut6.ButtonB := FALSE;
   BenchUut6.ButtonC := FALSE;
   TraceIn_Mode[75] := BenchUut6.Mode;
   TraceIn_ForwardButton[75] := BenchUut6.ForwardButton;
   TraceIn_ReverseButton[75] := BenchUut6.ReverseButton;
   TraceIn_SensorA[75] := BenchUut6.SensorA;
   TraceIn_SensorB[75] := BenchUut6.SensorB;
   TraceIn_SensorC[75] := BenchUut6.SensorC;
   TraceIn_ButtonA[75] := BenchUut6.ButtonA;
   TraceIn_ButtonB[75] := BenchUut6.ButtonB;
   TraceIn_ButtonC[75] := BenchUut6.ButtonC;
   BenchUut6();
   TraceOut_MotorForward[75] := BenchUut6.MotorForward;
   TraceOut_MotorReverse[75] := BenchUut6.MotorReverse;
   TraceOut_CompletionLight[75] := BenchUut6.CompletionLight;
   BenchCalls := BenchCalls + 1;
 76:
   BenchUut7.Mode := TRUE;
   BenchUut7.ForwardButton := FALSE;
   BenchUut7.ReverseButton := FALSE;
   BenchUut7.SensorA := FALSE;
   BenchUut7.SensorB := FALSE;
   BenchUut7.SensorC := FALSE;
   BenchUut7.ButtonA := FALSE;
   BenchUut7.ButtonB := TRUE;
   BenchUut7.ButtonC := TRUE;
   TraceIn_Mode[76] := BenchUut7.Mode;
   TraceIn_ForwardButton[76] := BenchUut7.ForwardButton;
   TraceIn_ReverseButton[76] := BenchUut7.ReverseButton;
   TraceIn_SensorA[76] := BenchUut7.SensorA;
   TraceIn_SensorB[76] := BenchUut7.SensorB;
   TraceIn_SensorC[76] := BenchUut7.SensorC;
   TraceIn_ButtonA[76] := BenchUut7.ButtonA;
   TraceIn_ButtonB[76] := BenchUut7.ButtonB;
   TraceIn_ButtonC[76] := BenchUut7.ButtonC;
   BenchUut7();
   TraceOut_MotorForward[76] := BenchUut7.MotorForward;
   TraceOut_MotorReverse[76] := BenchUut7.MotorReverse;
   TraceOut_CompletionLight[76] := BenchUut7.CompletionLight;
   BenchCalls := BenchCalls + 1;
 77:
   BenchUut7.Mode := TRUE;
   BenchUut7.ForwardButton := FALSE;
   BenchUut7.ReverseButton := FALSE;
   BenchUut7.SensorA := FALSE;
   BenchUut7.SensorB := FALSE;
   BenchUut7.SensorC := FALSE;
   BenchUut7.ButtonA := FALSE;
   BenchUut7.ButtonB := TRUE;
   BenchUut7.ButtonC := TRUE;
   TraceIn_Mode[77] := BenchUut7.Mode;
   TraceIn_ForwardButton[77] := BenchUut7.ForwardButton;
   TraceIn_ReverseButton[77] := BenchUut7.ReverseButton;
   TraceIn_SensorA[77] := BenchUut7.SensorA;
   TraceIn_SensorB[77] := BenchUut7.SensorB;
   TraceIn_SensorC[77] := BenchUut7.SensorC;
   TraceIn_ButtonA[77] := BenchUut7.ButtonA;
   TraceIn_ButtonB[77] := BenchUut7.ButtonB;
   TraceIn_ButtonC[77] := BenchUut7.ButtonC;
   BenchUut7();
   TraceOut_MotorForward[77] := BenchUut7.MotorForward;
   TraceOut_MotorReverse[77] := BenchUut7.MotorReverse;
   TraceOut_CompletionLight[77] := BenchUut7.CompletionLight;
   BenchCalls := BenchCalls + 1;
 78:
   BenchUut7.Mode := TRUE;
   BenchUut7.ForwardButton := FALSE;
   BenchUut7.ReverseButton := FALSE;
   BenchUut7.SensorA := FALSE;
   BenchUut7.SensorB := FALSE;
   BenchUut7.SensorC := FALSE;
   BenchUut7.ButtonA := FALSE;
   BenchUut7.ButtonB := TRUE;
   BenchUut7.ButtonC := TRUE;
   TraceIn_Mode[78] := BenchUut7.Mode;
   TraceIn_ForwardButton[78] := BenchUut7.ForwardButton;
   TraceIn_ReverseButton[78] := BenchUut7.ReverseButton;
   TraceIn_SensorA[78] := BenchUut7.SensorA;
   TraceIn_SensorB[78] := BenchUut7.SensorB;
   TraceIn_SensorC[78] := BenchUut7.SensorC;
   TraceIn_ButtonA[78] := BenchUut7.ButtonA;
   TraceIn_ButtonB[78] := BenchUut7.ButtonB;
   TraceIn_ButtonC[78] := BenchUut7.ButtonC;
   BenchUut7();
   TraceOut_MotorForward[78] := BenchUut7.MotorForward;
   TraceOut_MotorReverse[78] := BenchUut7.MotorReverse;
   TraceOut_CompletionLight[78] := BenchUut7.CompletionLight;
   BenchCalls := BenchCalls + 1;
 79:
   BenchUut7.Mode := TRUE;
   BenchUut7.ForwardButton := FALSE;
   BenchUut7.ReverseButton := FALSE;
   BenchUut7.SensorA := TRUE;
   BenchUut7.SensorB := FALSE;
   BenchUut7.SensorC := FALSE;
   BenchUut7.ButtonA := FALSE;
   BenchUut7.ButtonB := TRUE;
   BenchUut7.ButtonC := FALSE;
   TraceIn_Mode[79] := BenchUut7.Mode;
   TraceIn_ForwardButton[79] := BenchUut7.ForwardButton;
   TraceIn_ReverseButton[79] := BenchUut7.ReverseButton;
   TraceIn_SensorA[79] := BenchUut7.SensorA;
   TraceIn_SensorB[79] := BenchUut7.SensorB;
   TraceIn_SensorC[79] := BenchUut7.SensorC;
   TraceIn_ButtonA[79] := BenchUut7.ButtonA;
   TraceIn_ButtonB[79] := BenchUut7.ButtonB;
   TraceIn_ButtonC[79] := BenchUut7.ButtonC;
   BenchUut7();
   TraceOut_MotorForward[79] := BenchUut7.MotorForward;
   TraceOut_MotorReverse[79] := BenchUut7.MotorReverse;
   TraceOut_CompletionLight[79] := BenchUut7.CompletionLight;
   BenchCalls := BenchCalls + 1;
 80:
   BenchUut7.Mode := TRUE;
   BenchUut7.ForwardButton := FALSE;
   BenchUut7.ReverseButton := FALSE;
   BenchUut7.SensorA := TRUE;
   BenchUut7.SensorB := FALSE;
   BenchUut7.SensorC := FALSE;
   BenchUut7.ButtonA := FALSE;
   BenchUut7.ButtonB := TRUE;
   BenchUut7.ButtonC := FALSE;
   TraceIn_Mode[80] := BenchUut7.Mode;
   TraceIn_ForwardButton[80] := BenchUut7.ForwardButton;
   TraceIn_ReverseButton[80] := BenchUut7.ReverseButton;
   TraceIn_SensorA[80] := BenchUut7.SensorA;
   TraceIn_SensorB[80] := BenchUut7.SensorB;
   TraceIn_SensorC[80] := BenchUut7.SensorC;
   TraceIn_ButtonA[80] := BenchUut7.ButtonA;
   TraceIn_ButtonB[80] := BenchUut7.ButtonB;
   TraceIn_ButtonC[80] := BenchUut7.ButtonC;
   BenchUut7();
   TraceOut_MotorForward[80] := BenchUut7.MotorForward;
   TraceOut_MotorReverse[80] := BenchUut7.MotorReverse;
   TraceOut_CompletionLight[80] := BenchUut7.CompletionLight;
   BenchCalls := BenchCalls + 1;
 81:
   BenchUut7.Mode := TRUE;
   BenchUut7.ForwardButton := FALSE;
   BenchUut7.ReverseButton := FALSE;
   BenchUut7.SensorA := TRUE;
   BenchUut7.SensorB := FALSE;
   BenchUut7.SensorC := FALSE;
   BenchUut7.ButtonA := FALSE;
   BenchUut7.ButtonB := TRUE;
   BenchUut7.ButtonC := FALSE;
   TraceIn_Mode[81] := BenchUut7.Mode;
   TraceIn_ForwardButton[81] := BenchUut7.ForwardButton;
   TraceIn_ReverseButton[81] := BenchUut7.ReverseButton;
   TraceIn_SensorA[81] := BenchUut7.SensorA;
   TraceIn_SensorB[81] := BenchUut7.SensorB;
   TraceIn_SensorC[81] := BenchUut7.SensorC;
   TraceIn_ButtonA[81] := BenchUut7.ButtonA;
   TraceIn_ButtonB[81] := BenchUut7.ButtonB;
   TraceIn_ButtonC[81] := BenchUut7.ButtonC;
   BenchUut7();
   TraceOut_MotorForward[81] := BenchUut7.MotorForward;
   TraceOut_MotorReverse[81] := BenchUut7.MotorReverse;
   TraceOut_CompletionLight[81] := BenchUut7.CompletionLight;
   BenchCalls := BenchCalls + 1;
 END_CASE;
 BenchStep := BenchStep + 1;
 IF BenchStep >= 82 THEN BenchDone := TRUE; END_IF;
END_IF;
END_PROGRAM
